(* IEC 61131-3 sources: IEC61131-3_ST_SCL_Mutation_Generator/Tests/mutatedCodeGenbit, 69 files *)

(* ---- M001.st ---- *)
FUNCTION_BLOCK GEN_BIT
  VAR_INPUT
    IN0 : DWORD;
    IN1 : DWORD;
    IN2 : DWORD;
    IN3 : DWORD;
    CLK : BOOL;
    STEPS : INT;
    REP : INT;
    RST : BOOL;
  END_VAR
  VAR_OUTPUT
    Q0 : BOOL;
    Q1 : BOOL;
    Q2 : BOOL;
    Q3 : BOOL;
    CNT : INT;
    RUN : BOOL;
  END_VAR
  VAR
    r0 : DWORD;
    r1 : DWORD;
    r2 : DWORD;
    r3 : DWORD;
    rx : INT := 1;
  END_VAR

  (* check if number of runs is finished or rep <> 0 which means continuous *) (* MUTATED: REL_OP_REPLACE *)

  IF clk AND NOT rst THEN
  	run := (rep = 0) OR (rx <= rep);
  	IF run THEN
  		(* check for step counter reached and reset to 0 if cnt = steps *)
  		IF cnt = steps THEN
  			cnt := 0;
  		END_IF;

  		(* when cnt = 0 then reload the inputs into the registers *)
  		IF cnt = 0 THEN
  			r0 := in0;
  			r1 := in1;
  			r2 := in2;
  			r3 := in3;
  		END_IF;

  		(* when cnt < steps, shift the lowest bits to the outputs *)
  		IF (cnt < steps) THEN
              Q0 := BIT_OF_DWORD(r0,0); (* Q0 := r0.X0; *)
              Q1 := BIT_OF_DWORD(r1,0); (* Q1 := r1.X0; *)
              Q2 := BIT_OF_DWORD(r2,0); (* Q2 := r2.X0; *)
              Q3 := BIT_OF_DWORD(r3,0); (* Q3 := r3.X0; *)
  			r0 := SHR(r0,1);
  			r1 := SHR(r1,1);
  			r2 := SHR(r2,1);
  			r3 := SHR(r3,1);
  		END_IF;

  		(* increment the step counter *)
  		cnt := cnt +1;
  		IF (cnt = steps) AND (rep <> 0) THEN rx := rx +1; END_IF;
  		IF (rx > rep) AND (rep <> 0) THEN run := FALSE; END_IF;
  	END_IF;
  ELSE
  	IF rst THEN
  		run := FALSE;
  		Q0 := FALSE;
  		Q1 := FALSE;
  		Q2 := FALSE;
  		Q3 := FALSE;
  		r0 := DWORD#0;
  		r1 := DWORD#0;
  		r2 := DWORD#0;
  		r3 := DWORD#0;
  		cnt := 0;
  		rx := 1;
  	END_IF;
  END_IF;

  (*From OSCAT Library, www.oscat.de *)
END_FUNCTION_BLOCK

(* ---- M002.st ---- *)
FUNCTION_BLOCK GEN_BIT
  VAR_INPUT
    IN0 : DWORD;
    IN1 : DWORD;
    IN2 : DWORD;
    IN3 : DWORD;
    CLK : BOOL;
    STEPS : INT;
    REP : INT;
    RST : BOOL;
  END_VAR
  VAR_OUTPUT
    Q0 : BOOL;
    Q1 : BOOL;
    Q2 : BOOL;
    Q3 : BOOL;
    CNT : INT;
    RUN : BOOL;
  END_VAR
  VAR
    r0 : DWORD;
    r1 : DWORD;
    r2 : DWORD;
    r3 : DWORD;
    rx : INT := 1;
  END_VAR

  (* check if number of runs is finished or rep = 0 which means continuous *)

  IF clk AND NOT rst THEN
  	run := (rep <> 0) OR (rx <= rep); (* MUTATED: REL_OP_REPLACE *)
  	IF run THEN
  		(* check for step counter reached and reset to 0 if cnt = steps *)
  		IF cnt = steps THEN
  			cnt := 0;
  		END_IF;

  		(* when cnt = 0 then reload the inputs into the registers *)
  		IF cnt = 0 THEN
  			r0 := in0;
  			r1 := in1;
  			r2 := in2;
  			r3 := in3;
  		END_IF;

  		(* when cnt < steps, shift the lowest bits to the outputs *)
  		IF (cnt < steps) THEN
              Q0 := BIT_OF_DWORD(r0,0); (* Q0 := r0.X0; *)
              Q1 := BIT_OF_DWORD(r1,0); (* Q1 := r1.X0; *)
              Q2 := BIT_OF_DWORD(r2,0); (* Q2 := r2.X0; *)
              Q3 := BIT_OF_DWORD(r3,0); (* Q3 := r3.X0; *)
  			r0 := SHR(r0,1);
  			r1 := SHR(r1,1);
  			r2 := SHR(r2,1);
  			r3 := SHR(r3,1);
  		END_IF;

  		(* increment the step counter *)
  		cnt := cnt +1;
  		IF (cnt = steps) AND (rep <> 0) THEN rx := rx +1; END_IF;
  		IF (rx > rep) AND (rep <> 0) THEN run := FALSE; END_IF;
  	END_IF;
  ELSE
  	IF rst THEN
  		run := FALSE;
  		Q0 := FALSE;
  		Q1 := FALSE;
  		Q2 := FALSE;
  		Q3 := FALSE;
  		r0 := DWORD#0;
  		r1 := DWORD#0;
  		r2 := DWORD#0;
  		r3 := DWORD#0;
  		cnt := 0;
  		rx := 1;
  	END_IF;
  END_IF;

  (*From OSCAT Library, www.oscat.de *)
END_FUNCTION_BLOCK

(* ---- M003.st ---- *)
FUNCTION_BLOCK GEN_BIT
  VAR_INPUT
    IN0 : DWORD;
    IN1 : DWORD;
    IN2 : DWORD;
    IN3 : DWORD;
    CLK : BOOL;
    STEPS : INT;
    REP : INT;
    RST : BOOL;
  END_VAR
  VAR_OUTPUT
    Q0 : BOOL;
    Q1 : BOOL;
    Q2 : BOOL;
    Q3 : BOOL;
    CNT : INT;
    RUN : BOOL;
  END_VAR
  VAR
    r0 : DWORD;
    r1 : DWORD;
    r2 : DWORD;
    r3 : DWORD;
    rx : INT := 1;
  END_VAR

  (* check if number of runs is finished or rep = 0 which means continuous *)

  IF clk AND NOT rst THEN
  	run := (rep = 0) OR (rx >= rep); (* MUTATED: REL_OP_REPLACE *)
  	IF run THEN
  		(* check for step counter reached and reset to 0 if cnt = steps *)
  		IF cnt = steps THEN
  			cnt := 0;
  		END_IF;

  		(* when cnt = 0 then reload the inputs into the registers *)
  		IF cnt = 0 THEN
  			r0 := in0;
  			r1 := in1;
  			r2 := in2;
  			r3 := in3;
  		END_IF;

  		(* when cnt < steps, shift the lowest bits to the outputs *)
  		IF (cnt < steps) THEN
              Q0 := BIT_OF_DWORD(r0,0); (* Q0 := r0.X0; *)
              Q1 := BIT_OF_DWORD(r1,0); (* Q1 := r1.X0; *)
              Q2 := BIT_OF_DWORD(r2,0); (* Q2 := r2.X0; *)
              Q3 := BIT_OF_DWORD(r3,0); (* Q3 := r3.X0; *)
  			r0 := SHR(r0,1);
  			r1 := SHR(r1,1);
  			r2 := SHR(r2,1);
  			r3 := SHR(r3,1);
  		END_IF;

  		(* increment the step counter *)
  		cnt := cnt +1;
  		IF (cnt = steps) AND (rep <> 0) THEN rx := rx +1; END_IF;
  		IF (rx > rep) AND (rep <> 0) THEN run := FALSE; END_IF;
  	END_IF;
  ELSE
  	IF rst THEN
  		run := FALSE;
  		Q0 := FALSE;
  		Q1 := FALSE;
  		Q2 := FALSE;
  		Q3 := FALSE;
  		r0 := DWORD#0;
  		r1 := DWORD#0;
  		r2 := DWORD#0;
  		r3 := DWORD#0;
  		cnt := 0;
  		rx := 1;
  	END_IF;
  END_IF;

  (*From OSCAT Library, www.oscat.de *)
END_FUNCTION_BLOCK

(* ---- M004.st ---- *)
FUNCTION_BLOCK GEN_BIT
  VAR_INPUT
    IN0 : DWORD;
    IN1 : DWORD;
    IN2 : DWORD;
    IN3 : DWORD;
    CLK : BOOL;
    STEPS : INT;
    REP : INT;
    RST : BOOL;
  END_VAR
  VAR_OUTPUT
    Q0 : BOOL;
    Q1 : BOOL;
    Q2 : BOOL;
    Q3 : BOOL;
    CNT : INT;
    RUN : BOOL;
  END_VAR
  VAR
    r0 : DWORD;
    r1 : DWORD;
    r2 : DWORD;
    r3 : DWORD;
    rx : INT := 1;
  END_VAR

  (* check if number of runs is finished or rep = 0 which means continuous *)

  IF clk AND NOT rst THEN
  	run := (rep = 0) OR (rx <= rep);
  	IF run THEN
  		(* check for step counter reached and reset to 0 if cnt <> steps *) (* MUTATED: REL_OP_REPLACE *)
  		IF cnt = steps THEN
  			cnt := 0;
  		END_IF;

  		(* when cnt = 0 then reload the inputs into the registers *)
  		IF cnt = 0 THEN
  			r0 := in0;
  			r1 := in1;
  			r2 := in2;
  			r3 := in3;
  		END_IF;

  		(* when cnt < steps, shift the lowest bits to the outputs *)
  		IF (cnt < steps) THEN
              Q0 := BIT_OF_DWORD(r0,0); (* Q0 := r0.X0; *)
              Q1 := BIT_OF_DWORD(r1,0); (* Q1 := r1.X0; *)
              Q2 := BIT_OF_DWORD(r2,0); (* Q2 := r2.X0; *)
              Q3 := BIT_OF_DWORD(r3,0); (* Q3 := r3.X0; *)
  			r0 := SHR(r0,1);
  			r1 := SHR(r1,1);
  			r2 := SHR(r2,1);
  			r3 := SHR(r3,1);
  		END_IF;

  		(* increment the step counter *)
  		cnt := cnt +1;
  		IF (cnt = steps) AND (rep <> 0) THEN rx := rx +1; END_IF;
  		IF (rx > rep) AND (rep <> 0) THEN run := FALSE; END_IF;
  	END_IF;
  ELSE
  	IF rst THEN
  		run := FALSE;
  		Q0 := FALSE;
  		Q1 := FALSE;
  		Q2 := FALSE;
  		Q3 := FALSE;
  		r0 := DWORD#0;
  		r1 := DWORD#0;
  		r2 := DWORD#0;
  		r3 := DWORD#0;
  		cnt := 0;
  		rx := 1;
  	END_IF;
  END_IF;

  (*From OSCAT Library, www.oscat.de *)
END_FUNCTION_BLOCK

(* ---- M005.st ---- *)
FUNCTION_BLOCK GEN_BIT
  VAR_INPUT
    IN0 : DWORD;
    IN1 : DWORD;
    IN2 : DWORD;
    IN3 : DWORD;
    CLK : BOOL;
    STEPS : INT;
    REP : INT;
    RST : BOOL;
  END_VAR
  VAR_OUTPUT
    Q0 : BOOL;
    Q1 : BOOL;
    Q2 : BOOL;
    Q3 : BOOL;
    CNT : INT;
    RUN : BOOL;
  END_VAR
  VAR
    r0 : DWORD;
    r1 : DWORD;
    r2 : DWORD;
    r3 : DWORD;
    rx : INT := 1;
  END_VAR

  (* check if number of runs is finished or rep = 0 which means continuous *)

  IF clk AND NOT rst THEN
  	run := (rep = 0) OR (rx <= rep);
  	IF run THEN
  		(* check for step counter reached and reset to 0 if cnt = steps *)
  		IF cnt <> steps THEN (* MUTATED: REL_OP_REPLACE *)
  			cnt := 0;
  		END_IF;

  		(* when cnt = 0 then reload the inputs into the registers *)
  		IF cnt = 0 THEN
  			r0 := in0;
  			r1 := in1;
  			r2 := in2;
  			r3 := in3;
  		END_IF;

  		(* when cnt < steps, shift the lowest bits to the outputs *)
  		IF (cnt < steps) THEN
              Q0 := BIT_OF_DWORD(r0,0); (* Q0 := r0.X0; *)
              Q1 := BIT_OF_DWORD(r1,0); (* Q1 := r1.X0; *)
              Q2 := BIT_OF_DWORD(r2,0); (* Q2 := r2.X0; *)
              Q3 := BIT_OF_DWORD(r3,0); (* Q3 := r3.X0; *)
  			r0 := SHR(r0,1);
  			r1 := SHR(r1,1);
  			r2 := SHR(r2,1);
  			r3 := SHR(r3,1);
  		END_IF;

  		(* increment the step counter *)
  		cnt := cnt +1;
  		IF (cnt = steps) AND (rep <> 0) THEN rx := rx +1; END_IF;
  		IF (rx > rep) AND (rep <> 0) THEN run := FALSE; END_IF;
  	END_IF;
  ELSE
  	IF rst THEN
  		run := FALSE;
  		Q0 := FALSE;
  		Q1 := FALSE;
  		Q2 := FALSE;
  		Q3 := FALSE;
  		r0 := DWORD#0;
  		r1 := DWORD#0;
  		r2 := DWORD#0;
  		r3 := DWORD#0;
  		cnt := 0;
  		rx := 1;
  	END_IF;
  END_IF;

  (*From OSCAT Library, www.oscat.de *)
END_FUNCTION_BLOCK

(* ---- M006.st ---- *)
FUNCTION_BLOCK GEN_BIT
  VAR_INPUT
    IN0 : DWORD;
    IN1 : DWORD;
    IN2 : DWORD;
    IN3 : DWORD;
    CLK : BOOL;
    STEPS : INT;
    REP : INT;
    RST : BOOL;
  END_VAR
  VAR_OUTPUT
    Q0 : BOOL;
    Q1 : BOOL;
    Q2 : BOOL;
    Q3 : BOOL;
    CNT : INT;
    RUN : BOOL;
  END_VAR
  VAR
    r0 : DWORD;
    r1 : DWORD;
    r2 : DWORD;
    r3 : DWORD;
    rx : INT := 1;
  END_VAR

  (* check if number of runs is finished or rep = 0 which means continuous *)

  IF clk AND NOT rst THEN
  	run := (rep = 0) OR (rx <= rep);
  	IF run THEN
  		(* check for step counter reached and reset to 0 if cnt = steps *)
  		IF cnt = steps THEN
  			cnt := 0;
  		END_IF;

  		(* when cnt <> 0 then reload the inputs into the registers *) (* MUTATED: REL_OP_REPLACE *)
  		IF cnt = 0 THEN
  			r0 := in0;
  			r1 := in1;
  			r2 := in2;
  			r3 := in3;
  		END_IF;

  		(* when cnt < steps, shift the lowest bits to the outputs *)
  		IF (cnt < steps) THEN
              Q0 := BIT_OF_DWORD(r0,0); (* Q0 := r0.X0; *)
              Q1 := BIT_OF_DWORD(r1,0); (* Q1 := r1.X0; *)
              Q2 := BIT_OF_DWORD(r2,0); (* Q2 := r2.X0; *)
              Q3 := BIT_OF_DWORD(r3,0); (* Q3 := r3.X0; *)
  			r0 := SHR(r0,1);
  			r1 := SHR(r1,1);
  			r2 := SHR(r2,1);
  			r3 := SHR(r3,1);
  		END_IF;

  		(* increment the step counter *)
  		cnt := cnt +1;
  		IF (cnt = steps) AND (rep <> 0) THEN rx := rx +1; END_IF;
  		IF (rx > rep) AND (rep <> 0) THEN run := FALSE; END_IF;
  	END_IF;
  ELSE
  	IF rst THEN
  		run := FALSE;
  		Q0 := FALSE;
  		Q1 := FALSE;
  		Q2 := FALSE;
  		Q3 := FALSE;
  		r0 := DWORD#0;
  		r1 := DWORD#0;
  		r2 := DWORD#0;
  		r3 := DWORD#0;
  		cnt := 0;
  		rx := 1;
  	END_IF;
  END_IF;

  (*From OSCAT Library, www.oscat.de *)
END_FUNCTION_BLOCK

(* ---- M007.st ---- *)
FUNCTION_BLOCK GEN_BIT
  VAR_INPUT
    IN0 : DWORD;
    IN1 : DWORD;
    IN2 : DWORD;
    IN3 : DWORD;
    CLK : BOOL;
    STEPS : INT;
    REP : INT;
    RST : BOOL;
  END_VAR
  VAR_OUTPUT
    Q0 : BOOL;
    Q1 : BOOL;
    Q2 : BOOL;
    Q3 : BOOL;
    CNT : INT;
    RUN : BOOL;
  END_VAR
  VAR
    r0 : DWORD;
    r1 : DWORD;
    r2 : DWORD;
    r3 : DWORD;
    rx : INT := 1;
  END_VAR

  (* check if number of runs is finished or rep = 0 which means continuous *)

  IF clk AND NOT rst THEN
  	run := (rep = 0) OR (rx <= rep);
  	IF run THEN
  		(* check for step counter reached and reset to 0 if cnt = steps *)
  		IF cnt = steps THEN
  			cnt := 0;
  		END_IF;

  		(* when cnt = 0 then reload the inputs into the registers *)
  		IF cnt <> 0 THEN (* MUTATED: REL_OP_REPLACE *)
  			r0 := in0;
  			r1 := in1;
  			r2 := in2;
  			r3 := in3;
  		END_IF;

  		(* when cnt < steps, shift the lowest bits to the outputs *)
  		IF (cnt < steps) THEN
              Q0 := BIT_OF_DWORD(r0,0); (* Q0 := r0.X0; *)
              Q1 := BIT_OF_DWORD(r1,0); (* Q1 := r1.X0; *)
              Q2 := BIT_OF_DWORD(r2,0); (* Q2 := r2.X0; *)
              Q3 := BIT_OF_DWORD(r3,0); (* Q3 := r3.X0; *)
  			r0 := SHR(r0,1);
  			r1 := SHR(r1,1);
  			r2 := SHR(r2,1);
  			r3 := SHR(r3,1);
  		END_IF;

  		(* increment the step counter *)
  		cnt := cnt +1;
  		IF (cnt = steps) AND (rep <> 0) THEN rx := rx +1; END_IF;
  		IF (rx > rep) AND (rep <> 0) THEN run := FALSE; END_IF;
  	END_IF;
  ELSE
  	IF rst THEN
  		run := FALSE;
  		Q0 := FALSE;
  		Q1 := FALSE;
  		Q2 := FALSE;
  		Q3 := FALSE;
  		r0 := DWORD#0;
  		r1 := DWORD#0;
  		r2 := DWORD#0;
  		r3 := DWORD#0;
  		cnt := 0;
  		rx := 1;
  	END_IF;
  END_IF;

  (*From OSCAT Library, www.oscat.de *)
END_FUNCTION_BLOCK

(* ---- M008.st ---- *)
FUNCTION_BLOCK GEN_BIT
  VAR_INPUT
    IN0 : DWORD;
    IN1 : DWORD;
    IN2 : DWORD;
    IN3 : DWORD;
    CLK : BOOL;
    STEPS : INT;
    REP : INT;
    RST : BOOL;
  END_VAR
  VAR_OUTPUT
    Q0 : BOOL;
    Q1 : BOOL;
    Q2 : BOOL;
    Q3 : BOOL;
    CNT : INT;
    RUN : BOOL;
  END_VAR
  VAR
    r0 : DWORD;
    r1 : DWORD;
    r2 : DWORD;
    r3 : DWORD;
    rx : INT := 1;
  END_VAR

  (* check if number of runs is finished or rep = 0 which means continuous *)

  IF clk AND NOT rst THEN
  	run := (rep = 0) OR (rx <= rep);
  	IF run THEN
  		(* check for step counter reached and reset to 0 if cnt = steps *)
  		IF cnt = steps THEN
  			cnt := 0;
  		END_IF;

  		(* when cnt = 0 then reload the inputs into the registers *)
  		IF cnt = 0 THEN
  			r0 := in0;
  			r1 := in1;
  			r2 := in2;
  			r3 := in3;
  		END_IF;

  		(* when cnt > steps, shift the lowest bits to the outputs *) (* MUTATED: REL_OP_REPLACE *)
  		IF (cnt < steps) THEN
              Q0 := BIT_OF_DWORD(r0,0); (* Q0 := r0.X0; *)
              Q1 := BIT_OF_DWORD(r1,0); (* Q1 := r1.X0; *)
              Q2 := BIT_OF_DWORD(r2,0); (* Q2 := r2.X0; *)
              Q3 := BIT_OF_DWORD(r3,0); (* Q3 := r3.X0; *)
  			r0 := SHR(r0,1);
  			r1 := SHR(r1,1);
  			r2 := SHR(r2,1);
  			r3 := SHR(r3,1);
  		END_IF;

  		(* increment the step counter *)
  		cnt := cnt +1;
  		IF (cnt = steps) AND (rep <> 0) THEN rx := rx +1; END_IF;
  		IF (rx > rep) AND (rep <> 0) THEN run := FALSE; END_IF;
  	END_IF;
  ELSE
  	IF rst THEN
  		run := FALSE;
  		Q0 := FALSE;
  		Q1 := FALSE;
  		Q2 := FALSE;
  		Q3 := FALSE;
  		r0 := DWORD#0;
  		r1 := DWORD#0;
  		r2 := DWORD#0;
  		r3 := DWORD#0;
  		cnt := 0;
  		rx := 1;
  	END_IF;
  END_IF;

  (*From OSCAT Library, www.oscat.de *)
END_FUNCTION_BLOCK

(* ---- M009.st ---- *)
FUNCTION_BLOCK GEN_BIT
  VAR_INPUT
    IN0 : DWORD;
    IN1 : DWORD;
    IN2 : DWORD;
    IN3 : DWORD;
    CLK : BOOL;
    STEPS : INT;
    REP : INT;
    RST : BOOL;
  END_VAR
  VAR_OUTPUT
    Q0 : BOOL;
    Q1 : BOOL;
    Q2 : BOOL;
    Q3 : BOOL;
    CNT : INT;
    RUN : BOOL;
  END_VAR
  VAR
    r0 : DWORD;
    r1 : DWORD;
    r2 : DWORD;
    r3 : DWORD;
    rx : INT := 1;
  END_VAR

  (* check if number of runs is finished or rep = 0 which means continuous *)

  IF clk AND NOT rst THEN
  	run := (rep = 0) OR (rx <= rep);
  	IF run THEN
  		(* check for step counter reached and reset to 0 if cnt = steps *)
  		IF cnt = steps THEN
  			cnt := 0;
  		END_IF;

  		(* when cnt = 0 then reload the inputs into the registers *)
  		IF cnt = 0 THEN
  			r0 := in0;
  			r1 := in1;
  			r2 := in2;
  			r3 := in3;
  		END_IF;

  		(* when cnt < steps, shift the lowest bits to the outputs *)
  		IF (cnt > steps) THEN (* MUTATED: REL_OP_REPLACE *)
              Q0 := BIT_OF_DWORD(r0,0); (* Q0 := r0.X0; *)
              Q1 := BIT_OF_DWORD(r1,0); (* Q1 := r1.X0; *)
              Q2 := BIT_OF_DWORD(r2,0); (* Q2 := r2.X0; *)
              Q3 := BIT_OF_DWORD(r3,0); (* Q3 := r3.X0; *)
  			r0 := SHR(r0,1);
  			r1 := SHR(r1,1);
  			r2 := SHR(r2,1);
  			r3 := SHR(r3,1);
  		END_IF;

  		(* increment the step counter *)
  		cnt := cnt +1;
  		IF (cnt = steps) AND (rep <> 0) THEN rx := rx +1; END_IF;
  		IF (rx > rep) AND (rep <> 0) THEN run := FALSE; END_IF;
  	END_IF;
  ELSE
  	IF rst THEN
  		run := FALSE;
  		Q0 := FALSE;
  		Q1 := FALSE;
  		Q2 := FALSE;
  		Q3 := FALSE;
  		r0 := DWORD#0;
  		r1 := DWORD#0;
  		r2 := DWORD#0;
  		r3 := DWORD#0;
  		cnt := 0;
  		rx := 1;
  	END_IF;
  END_IF;

  (*From OSCAT Library, www.oscat.de *)
END_FUNCTION_BLOCK

(* ---- M010.st ---- *)
FUNCTION_BLOCK GEN_BIT
  VAR_INPUT
    IN0 : DWORD;
    IN1 : DWORD;
    IN2 : DWORD;
    IN3 : DWORD;
    CLK : BOOL;
    STEPS : INT;
    REP : INT;
    RST : BOOL;
  END_VAR
  VAR_OUTPUT
    Q0 : BOOL;
    Q1 : BOOL;
    Q2 : BOOL;
    Q3 : BOOL;
    CNT : INT;
    RUN : BOOL;
  END_VAR
  VAR
    r0 : DWORD;
    r1 : DWORD;
    r2 : DWORD;
    r3 : DWORD;
    rx : INT := 1;
  END_VAR

  (* check if number of runs is finished or rep = 0 which means continuous *)

  IF clk AND NOT rst THEN
  	run := (rep = 0) OR (rx <= rep);
  	IF run THEN
  		(* check for step counter reached and reset to 0 if cnt = steps *)
  		IF cnt = steps THEN
  			cnt := 0;
  		END_IF;

  		(* when cnt = 0 then reload the inputs into the registers *)
  		IF cnt = 0 THEN
  			r0 := in0;
  			r1 := in1;
  			r2 := in2;
  			r3 := in3;
  		END_IF;

  		(* when cnt < steps, shift the lowest bits to the outputs *)
  		IF (cnt < steps) THEN
              Q0 := BIT_OF_DWORD(r0,0); (* Q0 := r0.X0; *)
              Q1 := BIT_OF_DWORD(r1,0); (* Q1 := r1.X0; *)
              Q2 := BIT_OF_DWORD(r2,0); (* Q2 := r2.X0; *)
              Q3 := BIT_OF_DWORD(r3,0); (* Q3 := r3.X0; *)
  			r0 := SHR(r0,1);
  			r1 := SHR(r1,1);
  			r2 := SHR(r2,1);
  			r3 := SHR(r3,1);
  		END_IF;

  		(* increment the step counter *)
  		cnt := cnt +1;
  		IF (cnt <> steps) AND (rep <> 0) THEN rx := rx +1; END_IF; (* MUTATED: REL_OP_REPLACE *)
  		IF (rx > rep) AND (rep <> 0) THEN run := FALSE; END_IF;
  	END_IF;
  ELSE
  	IF rst THEN
  		run := FALSE;
  		Q0 := FALSE;
  		Q1 := FALSE;
  		Q2 := FALSE;
  		Q3 := FALSE;
  		r0 := DWORD#0;
  		r1 := DWORD#0;
  		r2 := DWORD#0;
  		r3 := DWORD#0;
  		cnt := 0;
  		rx := 1;
  	END_IF;
  END_IF;

  (*From OSCAT Library, www.oscat.de *)
END_FUNCTION_BLOCK

(* ---- M011.st ---- *)
FUNCTION_BLOCK GEN_BIT
  VAR_INPUT
    IN0 : DWORD;
    IN1 : DWORD;
    IN2 : DWORD;
    IN3 : DWORD;
    CLK : BOOL;
    STEPS : INT;
    REP : INT;
    RST : BOOL;
  END_VAR
  VAR_OUTPUT
    Q0 : BOOL;
    Q1 : BOOL;
    Q2 : BOOL;
    Q3 : BOOL;
    CNT : INT;
    RUN : BOOL;
  END_VAR
  VAR
    r0 : DWORD;
    r1 : DWORD;
    r2 : DWORD;
    r3 : DWORD;
    rx : INT := 1;
  END_VAR

  (* check if number of runs is finished or rep = 0 which means continuous *)

  IF clk AND NOT rst THEN
  	run := (rep = 0) OR (rx <= rep);
  	IF run THEN
  		(* check for step counter reached and reset to 0 if cnt = steps *)
  		IF cnt = steps THEN
  			cnt := 0;
  		END_IF;

  		(* when cnt = 0 then reload the inputs into the registers *)
  		IF cnt = 0 THEN
  			r0 := in0;
  			r1 := in1;
  			r2 := in2;
  			r3 := in3;
  		END_IF;

  		(* when cnt < steps, shift the lowest bits to the outputs *)
  		IF (cnt < steps) THEN
              Q0 := BIT_OF_DWORD(r0,0); (* Q0 := r0.X0; *)
              Q1 := BIT_OF_DWORD(r1,0); (* Q1 := r1.X0; *)
              Q2 := BIT_OF_DWORD(r2,0); (* Q2 := r2.X0; *)
              Q3 := BIT_OF_DWORD(r3,0); (* Q3 := r3.X0; *)
  			r0 := SHR(r0,1);
  			r1 := SHR(r1,1);
  			r2 := SHR(r2,1);
  			r3 := SHR(r3,1);
  		END_IF;

  		(* increment the step counter *)
  		cnt := cnt +1;
  		IF (cnt = steps) AND (rep = 0) THEN rx := rx +1; END_IF; (* MUTATED: REL_OP_REPLACE *)
  		IF (rx > rep) AND (rep <> 0) THEN run := FALSE; END_IF;
  	END_IF;
  ELSE
  	IF rst THEN
  		run := FALSE;
  		Q0 := FALSE;
  		Q1 := FALSE;
  		Q2 := FALSE;
  		Q3 := FALSE;
  		r0 := DWORD#0;
  		r1 := DWORD#0;
  		r2 := DWORD#0;
  		r3 := DWORD#0;
  		cnt := 0;
  		rx := 1;
  	END_IF;
  END_IF;

  (*From OSCAT Library, www.oscat.de *)
END_FUNCTION_BLOCK

(* ---- M012.st ---- *)
FUNCTION_BLOCK GEN_BIT
  VAR_INPUT
    IN0 : DWORD;
    IN1 : DWORD;
    IN2 : DWORD;
    IN3 : DWORD;
    CLK : BOOL;
    STEPS : INT;
    REP : INT;
    RST : BOOL;
  END_VAR
  VAR_OUTPUT
    Q0 : BOOL;
    Q1 : BOOL;
    Q2 : BOOL;
    Q3 : BOOL;
    CNT : INT;
    RUN : BOOL;
  END_VAR
  VAR
    r0 : DWORD;
    r1 : DWORD;
    r2 : DWORD;
    r3 : DWORD;
    rx : INT := 1;
  END_VAR

  (* check if number of runs is finished or rep = 0 which means continuous *)

  IF clk AND NOT rst THEN
  	run := (rep = 0) OR (rx <= rep);
  	IF run THEN
  		(* check for step counter reached and reset to 0 if cnt = steps *)
  		IF cnt = steps THEN
  			cnt := 0;
  		END_IF;

  		(* when cnt = 0 then reload the inputs into the registers *)
  		IF cnt = 0 THEN
  			r0 := in0;
  			r1 := in1;
  			r2 := in2;
  			r3 := in3;
  		END_IF;

  		(* when cnt < steps, shift the lowest bits to the outputs *)
  		IF (cnt < steps) THEN
              Q0 := BIT_OF_DWORD(r0,0); (* Q0 := r0.X0; *)
              Q1 := BIT_OF_DWORD(r1,0); (* Q1 := r1.X0; *)
              Q2 := BIT_OF_DWORD(r2,0); (* Q2 := r2.X0; *)
              Q3 := BIT_OF_DWORD(r3,0); (* Q3 := r3.X0; *)
  			r0 := SHR(r0,1);
  			r1 := SHR(r1,1);
  			r2 := SHR(r2,1);
  			r3 := SHR(r3,1);
  		END_IF;

  		(* increment the step counter *)
  		cnt := cnt +1;
  		IF (cnt = steps) AND (rep <> 0) THEN rx := rx +1; END_IF;
  		IF (rx < rep) AND (rep <> 0) THEN run := FALSE; END_IF; (* MUTATED: REL_OP_REPLACE *)
  	END_IF;
  ELSE
  	IF rst THEN
  		run := FALSE;
  		Q0 := FALSE;
  		Q1 := FALSE;
  		Q2 := FALSE;
  		Q3 := FALSE;
  		r0 := DWORD#0;
  		r1 := DWORD#0;
  		r2 := DWORD#0;
  		r3 := DWORD#0;
  		cnt := 0;
  		rx := 1;
  	END_IF;
  END_IF;

  (*From OSCAT Library, www.oscat.de *)
END_FUNCTION_BLOCK

(* ---- M013.st ---- *)
FUNCTION_BLOCK GEN_BIT
  VAR_INPUT
    IN0 : DWORD;
    IN1 : DWORD;
    IN2 : DWORD;
    IN3 : DWORD;
    CLK : BOOL;
    STEPS : INT;
    REP : INT;
    RST : BOOL;
  END_VAR
  VAR_OUTPUT
    Q0 : BOOL;
    Q1 : BOOL;
    Q2 : BOOL;
    Q3 : BOOL;
    CNT : INT;
    RUN : BOOL;
  END_VAR
  VAR
    r0 : DWORD;
    r1 : DWORD;
    r2 : DWORD;
    r3 : DWORD;
    rx : INT := 1;
  END_VAR

  (* check if number of runs is finished or rep = 0 which means continuous *)

  IF clk AND NOT rst THEN
  	run := (rep = 0) OR (rx <= rep);
  	IF run THEN
  		(* check for step counter reached and reset to 0 if cnt = steps *)
  		IF cnt = steps THEN
  			cnt := 0;
  		END_IF;

  		(* when cnt = 0 then reload the inputs into the registers *)
  		IF cnt = 0 THEN
  			r0 := in0;
  			r1 := in1;
  			r2 := in2;
  			r3 := in3;
  		END_IF;

  		(* when cnt < steps, shift the lowest bits to the outputs *)
  		IF (cnt < steps) THEN
              Q0 := BIT_OF_DWORD(r0,0); (* Q0 := r0.X0; *)
              Q1 := BIT_OF_DWORD(r1,0); (* Q1 := r1.X0; *)
              Q2 := BIT_OF_DWORD(r2,0); (* Q2 := r2.X0; *)
              Q3 := BIT_OF_DWORD(r3,0); (* Q3 := r3.X0; *)
  			r0 := SHR(r0,1);
  			r1 := SHR(r1,1);
  			r2 := SHR(r2,1);
  			r3 := SHR(r3,1);
  		END_IF;

  		(* increment the step counter *)
  		cnt := cnt +1;
  		IF (cnt = steps) AND (rep <> 0) THEN rx := rx +1; END_IF;
  		IF (rx > rep) AND (rep = 0) THEN run := FALSE; END_IF; (* MUTATED: REL_OP_REPLACE *)
  	END_IF;
  ELSE
  	IF rst THEN
  		run := FALSE;
  		Q0 := FALSE;
  		Q1 := FALSE;
  		Q2 := FALSE;
  		Q3 := FALSE;
  		r0 := DWORD#0;
  		r1 := DWORD#0;
  		r2 := DWORD#0;
  		r3 := DWORD#0;
  		cnt := 0;
  		rx := 1;
  	END_IF;
  END_IF;

  (*From OSCAT Library, www.oscat.de *)
END_FUNCTION_BLOCK

(* ---- M014.st ---- *)
FUNCTION_BLOCK GEN_BIT
  VAR_INPUT
    IN0 : DWORD;
    IN1 : DWORD;
    IN2 : DWORD;
    IN3 : DWORD;
    CLK : BOOL;
    STEPS : INT;
    REP : INT;
    RST : BOOL;
  END_VAR
  VAR_OUTPUT
    Q0 : BOOL;
    Q1 : BOOL;
    Q2 : BOOL;
    Q3 : BOOL;
    CNT : INT;
    RUN : BOOL;
  END_VAR
  VAR
    r0 : DWORD;
    r1 : DWORD;
    r2 : DWORD;
    r3 : DWORD;
    rx : INT := 1;
  END_VAR

  (* check if number of runs is finished or rep = 0 which means continuous *)

  IF clk OR NOT rst THEN (* MUTATED: LOGICAL_OP_REPLACE *)
  	run := (rep = 0) OR (rx <= rep);
  	IF run THEN
  		(* check for step counter reached and reset to 0 if cnt = steps *)
  		IF cnt = steps THEN
  			cnt := 0;
  		END_IF;

  		(* when cnt = 0 then reload the inputs into the registers *)
  		IF cnt = 0 THEN
  			r0 := in0;
  			r1 := in1;
  			r2 := in2;
  			r3 := in3;
  		END_IF;

  		(* when cnt < steps, shift the lowest bits to the outputs *)
  		IF (cnt < steps) THEN
              Q0 := BIT_OF_DWORD(r0,0); (* Q0 := r0.X0; *)
              Q1 := BIT_OF_DWORD(r1,0); (* Q1 := r1.X0; *)
              Q2 := BIT_OF_DWORD(r2,0); (* Q2 := r2.X0; *)
              Q3 := BIT_OF_DWORD(r3,0); (* Q3 := r3.X0; *)
  			r0 := SHR(r0,1);
  			r1 := SHR(r1,1);
  			r2 := SHR(r2,1);
  			r3 := SHR(r3,1);
  		END_IF;

  		(* increment the step counter *)
  		cnt := cnt +1;
  		IF (cnt = steps) AND (rep <> 0) THEN rx := rx +1; END_IF;
  		IF (rx > rep) AND (rep <> 0) THEN run := FALSE; END_IF;
  	END_IF;
  ELSE
  	IF rst THEN
  		run := FALSE;
  		Q0 := FALSE;
  		Q1 := FALSE;
  		Q2 := FALSE;
  		Q3 := FALSE;
  		r0 := DWORD#0;
  		r1 := DWORD#0;
  		r2 := DWORD#0;
  		r3 := DWORD#0;
  		cnt := 0;
  		rx := 1;
  	END_IF;
  END_IF;

  (*From OSCAT Library, www.oscat.de *)
END_FUNCTION_BLOCK

(* ---- M015.st ---- *)
FUNCTION_BLOCK GEN_BIT
  VAR_INPUT
    IN0 : DWORD;
    IN1 : DWORD;
    IN2 : DWORD;
    IN3 : DWORD;
    CLK : BOOL;
    STEPS : INT;
    REP : INT;
    RST : BOOL;
  END_VAR
  VAR_OUTPUT
    Q0 : BOOL;
    Q1 : BOOL;
    Q2 : BOOL;
    Q3 : BOOL;
    CNT : INT;
    RUN : BOOL;
  END_VAR
  VAR
    r0 : DWORD;
    r1 : DWORD;
    r2 : DWORD;
    r3 : DWORD;
    rx : INT := 1;
  END_VAR

  (* check if number of runs is finished or rep = 0 which means continuous *)

  IF clk AND NOT rst THEN
  	run := (rep = 0) AND (rx <= rep); (* MUTATED: LOGICAL_OP_REPLACE *)
  	IF run THEN
  		(* check for step counter reached and reset to 0 if cnt = steps *)
  		IF cnt = steps THEN
  			cnt := 0;
  		END_IF;

  		(* when cnt = 0 then reload the inputs into the registers *)
  		IF cnt = 0 THEN
  			r0 := in0;
  			r1 := in1;
  			r2 := in2;
  			r3 := in3;
  		END_IF;

  		(* when cnt < steps, shift the lowest bits to the outputs *)
  		IF (cnt < steps) THEN
              Q0 := BIT_OF_DWORD(r0,0); (* Q0 := r0.X0; *)
              Q1 := BIT_OF_DWORD(r1,0); (* Q1 := r1.X0; *)
              Q2 := BIT_OF_DWORD(r2,0); (* Q2 := r2.X0; *)
              Q3 := BIT_OF_DWORD(r3,0); (* Q3 := r3.X0; *)
  			r0 := SHR(r0,1);
  			r1 := SHR(r1,1);
  			r2 := SHR(r2,1);
  			r3 := SHR(r3,1);
  		END_IF;

  		(* increment the step counter *)
  		cnt := cnt +1;
  		IF (cnt = steps) AND (rep <> 0) THEN rx := rx +1; END_IF;
  		IF (rx > rep) AND (rep <> 0) THEN run := FALSE; END_IF;
  	END_IF;
  ELSE
  	IF rst THEN
  		run := FALSE;
  		Q0 := FALSE;
  		Q1 := FALSE;
  		Q2 := FALSE;
  		Q3 := FALSE;
  		r0 := DWORD#0;
  		r1 := DWORD#0;
  		r2 := DWORD#0;
  		r3 := DWORD#0;
  		cnt := 0;
  		rx := 1;
  	END_IF;
  END_IF;

  (*From OSCAT Library, www.oscat.de *)
END_FUNCTION_BLOCK

(* ---- M016.st ---- *)
FUNCTION_BLOCK GEN_BIT
  VAR_INPUT
    IN0 : DWORD;
    IN1 : DWORD;
    IN2 : DWORD;
    IN3 : DWORD;
    CLK : BOOL;
    STEPS : INT;
    REP : INT;
    RST : BOOL;
  END_VAR
  VAR_OUTPUT
    Q0 : BOOL;
    Q1 : BOOL;
    Q2 : BOOL;
    Q3 : BOOL;
    CNT : INT;
    RUN : BOOL;
  END_VAR
  VAR
    r0 : DWORD;
    r1 : DWORD;
    r2 : DWORD;
    r3 : DWORD;
    rx : INT := 1;
  END_VAR

  (* check if number of runs is finished or rep = 0 which means continuous *)

  IF clk AND NOT rst THEN
  	run := (rep = 0) OR (rx <= rep);
  	IF run THEN
  		(* check for step counter reached and reset to 0 if cnt = steps *)
  		IF cnt = steps THEN
  			cnt := 0;
  		END_IF;

  		(* when cnt = 0 then reload the inputs into the registers *)
  		IF cnt = 0 THEN
  			r0 := in0;
  			r1 := in1;
  			r2 := in2;
  			r3 := in3;
  		END_IF;

  		(* when cnt < steps, shift the lowest bits to the outputs *)
  		IF (cnt < steps) THEN
              Q0 := BIT_OF_DWORD(r0,0); (* Q0 := r0.X0; *)
              Q1 := BIT_OF_DWORD(r1,0); (* Q1 := r1.X0; *)
              Q2 := BIT_OF_DWORD(r2,0); (* Q2 := r2.X0; *)
              Q3 := BIT_OF_DWORD(r3,0); (* Q3 := r3.X0; *)
  			r0 := SHR(r0,1);
  			r1 := SHR(r1,1);
  			r2 := SHR(r2,1);
  			r3 := SHR(r3,1);
  		END_IF;

  		(* increment the step counter *)
  		cnt := cnt +1;
  		IF (cnt = steps) OR (rep <> 0) THEN rx := rx +1; END_IF; (* MUTATED: LOGICAL_OP_REPLACE *)
  		IF (rx > rep) AND (rep <> 0) THEN run := FALSE; END_IF;
  	END_IF;
  ELSE
  	IF rst THEN
  		run := FALSE;
  		Q0 := FALSE;
  		Q1 := FALSE;
  		Q2 := FALSE;
  		Q3 := FALSE;
  		r0 := DWORD#0;
  		r1 := DWORD#0;
  		r2 := DWORD#0;
  		r3 := DWORD#0;
  		cnt := 0;
  		rx := 1;
  	END_IF;
  END_IF;

  (*From OSCAT Library, www.oscat.de *)
END_FUNCTION_BLOCK

(* ---- M017.st ---- *)
FUNCTION_BLOCK GEN_BIT
  VAR_INPUT
    IN0 : DWORD;
    IN1 : DWORD;
    IN2 : DWORD;
    IN3 : DWORD;
    CLK : BOOL;
    STEPS : INT;
    REP : INT;
    RST : BOOL;
  END_VAR
  VAR_OUTPUT
    Q0 : BOOL;
    Q1 : BOOL;
    Q2 : BOOL;
    Q3 : BOOL;
    CNT : INT;
    RUN : BOOL;
  END_VAR
  VAR
    r0 : DWORD;
    r1 : DWORD;
    r2 : DWORD;
    r3 : DWORD;
    rx : INT := 1;
  END_VAR

  (* check if number of runs is finished or rep = 0 which means continuous *)

  IF clk AND NOT rst THEN
  	run := (rep = 0) OR (rx <= rep);
  	IF run THEN
  		(* check for step counter reached and reset to 0 if cnt = steps *)
  		IF cnt = steps THEN
  			cnt := 0;
  		END_IF;

  		(* when cnt = 0 then reload the inputs into the registers *)
  		IF cnt = 0 THEN
  			r0 := in0;
  			r1 := in1;
  			r2 := in2;
  			r3 := in3;
  		END_IF;

  		(* when cnt < steps, shift the lowest bits to the outputs *)
  		IF (cnt < steps) THEN
              Q0 := BIT_OF_DWORD(r0,0); (* Q0 := r0.X0; *)
              Q1 := BIT_OF_DWORD(r1,0); (* Q1 := r1.X0; *)
              Q2 := BIT_OF_DWORD(r2,0); (* Q2 := r2.X0; *)
              Q3 := BIT_OF_DWORD(r3,0); (* Q3 := r3.X0; *)
  			r0 := SHR(r0,1);
  			r1 := SHR(r1,1);
  			r2 := SHR(r2,1);
  			r3 := SHR(r3,1);
  		END_IF;

  		(* increment the step counter *)
  		cnt := cnt +1;
  		IF (cnt = steps) AND (rep <> 0) THEN rx := rx +1; END_IF;
  		IF (rx > rep) OR (rep <> 0) THEN run := FALSE; END_IF; (* MUTATED: LOGICAL_OP_REPLACE *)
  	END_IF;
  ELSE
  	IF rst THEN
  		run := FALSE;
  		Q0 := FALSE;
  		Q1 := FALSE;
  		Q2 := FALSE;
  		Q3 := FALSE;
  		r0 := DWORD#0;
  		r1 := DWORD#0;
  		r2 := DWORD#0;
  		r3 := DWORD#0;
  		cnt := 0;
  		rx := 1;
  	END_IF;
  END_IF;

  (*From OSCAT Library, www.oscat.de *)
END_FUNCTION_BLOCK

(* ---- M018.st ---- *)
FUNCTION_BLOCK GEN_BIT
  VAR_INPUT
    IN0 : DWORD;
    IN1 : DWORD;
    IN2 : DWORD;
    IN3 : DWORD;
    CLK : BOOL;
    STEPS : INT;
    REP : INT;
    RST : BOOL;
  END_VAR
  VAR_OUTPUT
    Q0 : BOOL;
    Q1 : BOOL;
    Q2 : BOOL;
    Q3 : BOOL;
    CNT : INT;
    RUN : BOOL;
  END_VAR
  VAR
    r0 : DWORD;
    r1 : DWORD;
    r2 : DWORD;
    r3 : DWORD;
    rx : INT := 1;
  END_VAR

  (* check if number of runs is finished or rep = 0 which means continuous *)

  IF clk AND NOT rst THEN
  	run := (rep = 0) OR (rx <= rep);
  	IF run THEN
  		(* check for step counter reached and reset to 0 if cnt = steps *)
  		IF cnt = steps THEN
  			cnt := 0;
  		END_IF;

  		(* when cnt = 0 then reload the inputs into the registers *)
  		IF cnt = 0 THEN
  			r0 := in0;
  			r1 := in1;
  			r2 := in2;
  			r3 := in3;
  		END_IF;

  		(* when cnt < steps, shift the lowest bits to the outputs *)
  		IF (cnt < steps) THEN
              Q0 := BIT_OF_DWORD(r0,0); (* Q0 := r0.X0; *)
              Q1 := BIT_OF_DWORD(r1,0); (* Q1 := r1.X0; *)
              Q2 := BIT_OF_DWORD(r2,0); (* Q2 := r2.X0; *)
              Q3 := BIT_OF_DWORD(r3,0); (* Q3 := r3.X0; *)
  			r0 := SHR(r0,1);
  			r1 := SHR(r1,1);
  			r2 := SHR(r2,1);
  			r3 := SHR(r3,1);
  		END_IF;

  		(* increment the step counter *)
  		cnt := cnt -1; (* MUTATED: ARITH_OP_REPLACE *)
  		IF (cnt = steps) AND (rep <> 0) THEN rx := rx +1; END_IF;
  		IF (rx > rep) AND (rep <> 0) THEN run := FALSE; END_IF;
  	END_IF;
  ELSE
  	IF rst THEN
  		run := FALSE;
  		Q0 := FALSE;
  		Q1 := FALSE;
  		Q2 := FALSE;
  		Q3 := FALSE;
  		r0 := DWORD#0;
  		r1 := DWORD#0;
  		r2 := DWORD#0;
  		r3 := DWORD#0;
  		cnt := 0;
  		rx := 1;
  	END_IF;
  END_IF;

  (*From OSCAT Library, www.oscat.de *)
END_FUNCTION_BLOCK

(* ---- M019.st ---- *)
FUNCTION_BLOCK GEN_BIT
  VAR_INPUT
    IN0 : DWORD;
    IN1 : DWORD;
    IN2 : DWORD;
    IN3 : DWORD;
    CLK : BOOL;
    STEPS : INT;
    REP : INT;
    RST : BOOL;
  END_VAR
  VAR_OUTPUT
    Q0 : BOOL;
    Q1 : BOOL;
    Q2 : BOOL;
    Q3 : BOOL;
    CNT : INT;
    RUN : BOOL;
  END_VAR
  VAR
    r0 : DWORD;
    r1 : DWORD;
    r2 : DWORD;
    r3 : DWORD;
    rx : INT := 1;
  END_VAR

  (* check if number of runs is finished or rep = 0 which means continuous *)

  IF clk AND NOT rst THEN
  	run := (rep = 0) OR (rx <= rep);
  	IF run THEN
  		(* check for step counter reached and reset to 0 if cnt = steps *)
  		IF cnt = steps THEN
  			cnt := 0;
  		END_IF;

  		(* when cnt = 0 then reload the inputs into the registers *)
  		IF cnt = 0 THEN
  			r0 := in0;
  			r1 := in1;
  			r2 := in2;
  			r3 := in3;
  		END_IF;

  		(* when cnt < steps, shift the lowest bits to the outputs *)
  		IF (cnt < steps) THEN
              Q0 := BIT_OF_DWORD(r0,0); (* Q0 := r0.X0; *)
              Q1 := BIT_OF_DWORD(r1,0); (* Q1 := r1.X0; *)
              Q2 := BIT_OF_DWORD(r2,0); (* Q2 := r2.X0; *)
              Q3 := BIT_OF_DWORD(r3,0); (* Q3 := r3.X0; *)
  			r0 := SHR(r0,1);
  			r1 := SHR(r1,1);
  			r2 := SHR(r2,1);
  			r3 := SHR(r3,1);
  		END_IF;

  		(* increment the step counter *)
  		cnt := cnt +1;
  		IF (cnt = steps) AND (rep <> 0) THEN rx := rx -1; END_IF; (* MUTATED: ARITH_OP_REPLACE *)
  		IF (rx > rep) AND (rep <> 0) THEN run := FALSE; END_IF;
  	END_IF;
  ELSE
  	IF rst THEN
  		run := FALSE;
  		Q0 := FALSE;
  		Q1 := FALSE;
  		Q2 := FALSE;
  		Q3 := FALSE;
  		r0 := DWORD#0;
  		r1 := DWORD#0;
  		r2 := DWORD#0;
  		r3 := DWORD#0;
  		cnt := 0;
  		rx := 1;
  	END_IF;
  END_IF;

  (*From OSCAT Library, www.oscat.de *)
END_FUNCTION_BLOCK

(* ---- M020.st ---- *)
FUNCTION_BLOCK GEN_BIT
  VAR_INPUT
    IN0 : DWORD;
    IN1 : DWORD;
    IN2 : DWORD;
    IN3 : DWORD;
    CLK : BOOL;
    STEPS : INT;
    REP : INT;
    RST : BOOL;
  END_VAR
  VAR_OUTPUT
    Q0 : BOOL;
    Q1 : BOOL;
    Q2 : BOOL;
    Q3 : BOOL;
    CNT : INT;
    RUN : BOOL;
  END_VAR
  VAR
    r0 : DWORD;
    r1 : DWORD;
    r2 : DWORD;
    r3 : DWORD;
    rx : INT := 1;
  END_VAR

  (* check if number of runs is finished or rep = 0 which means continuous *)

  IF clk AND NOT rst THEN
  	run := (rep = 0) OR (rx <= rep);
  	IF run THEN
  		(* check for step counter reached and reset to 0 if cnt = steps *)
  		IF cnt = steps THEN
  			cnt := 0;
  		END_IF;

  		(* when cnt = 0 then reload the inputs into the registers *)
  		IF cnt = 0 THEN
  			r0 := in0;
  			r1 := in1;
  			r2 := in2;
  			r3 := in3;
  		END_IF;

  		(* when cnt < steps, shift the lowest bits to the outputs *)
  		IF (cnt < steps) THEN
              Q0 := BIT_OF_DWORD(r0,0); (* Q0 := r0.X0; *)
              Q1 := BIT_OF_DWORD(r1,0); (* Q1 := r1.X0; *)
              Q2 := BIT_OF_DWORD(r2,0); (* Q2 := r2.X0; *)
              Q3 := BIT_OF_DWORD(r3,0); (* Q3 := r3.X0; *)
  			r0 := SHR(r0,1);
  			r1 := SHR(r1,1);
  			r2 := SHR(r2,1);
  			r3 := SHR(r3,1);
  		END_IF;

  		(* increment the step counter *)
  		cnt := cnt +1;
  		IF (cnt = steps) AND (rep <> 0) THEN rx := rx +1; END_IF;
  		IF (rx > rep) AND (rep <> 0) THEN run := TRUE; END_IF; (* MUTATED: BOOL_CONST_REPLACE *)
  	END_IF;
  ELSE
  	IF rst THEN
  		run := FALSE;
  		Q0 := FALSE;
  		Q1 := FALSE;
  		Q2 := FALSE;
  		Q3 := FALSE;
  		r0 := DWORD#0;
  		r1 := DWORD#0;
  		r2 := DWORD#0;
  		r3 := DWORD#0;
  		cnt := 0;
  		rx := 1;
  	END_IF;
  END_IF;

  (*From OSCAT Library, www.oscat.de *)
END_FUNCTION_BLOCK

(* ---- M021.st ---- *)
FUNCTION_BLOCK GEN_BIT
  VAR_INPUT
    IN0 : DWORD;
    IN1 : DWORD;
    IN2 : DWORD;
    IN3 : DWORD;
    CLK : BOOL;
    STEPS : INT;
    REP : INT;
    RST : BOOL;
  END_VAR
  VAR_OUTPUT
    Q0 : BOOL;
    Q1 : BOOL;
    Q2 : BOOL;
    Q3 : BOOL;
    CNT : INT;
    RUN : BOOL;
  END_VAR
  VAR
    r0 : DWORD;
    r1 : DWORD;
    r2 : DWORD;
    r3 : DWORD;
    rx : INT := 1;
  END_VAR

  (* check if number of runs is finished or rep = 0 which means continuous *)

  IF clk AND NOT rst THEN
  	run := (rep = 0) OR (rx <= rep);
  	IF run THEN
  		(* check for step counter reached and reset to 0 if cnt = steps *)
  		IF cnt = steps THEN
  			cnt := 0;
  		END_IF;

  		(* when cnt = 0 then reload the inputs into the registers *)
  		IF cnt = 0 THEN
  			r0 := in0;
  			r1 := in1;
  			r2 := in2;
  			r3 := in3;
  		END_IF;

  		(* when cnt < steps, shift the lowest bits to the outputs *)
  		IF (cnt < steps) THEN
              Q0 := BIT_OF_DWORD(r0,0); (* Q0 := r0.X0; *)
              Q1 := BIT_OF_DWORD(r1,0); (* Q1 := r1.X0; *)
              Q2 := BIT_OF_DWORD(r2,0); (* Q2 := r2.X0; *)
              Q3 := BIT_OF_DWORD(r3,0); (* Q3 := r3.X0; *)
  			r0 := SHR(r0,1);
  			r1 := SHR(r1,1);
  			r2 := SHR(r2,1);
  			r3 := SHR(r3,1);
  		END_IF;

  		(* increment the step counter *)
  		cnt := cnt +1;
  		IF (cnt = steps) AND (rep <> 0) THEN rx := rx +1; END_IF;
  		IF (rx > rep) AND (rep <> 0) THEN run := FALSE; END_IF;
  	END_IF;
  ELSE
  	IF rst THEN
  		run := TRUE; (* MUTATED: BOOL_CONST_REPLACE *)
  		Q0 := FALSE;
  		Q1 := FALSE;
  		Q2 := FALSE;
  		Q3 := FALSE;
  		r0 := DWORD#0;
  		r1 := DWORD#0;
  		r2 := DWORD#0;
  		r3 := DWORD#0;
  		cnt := 0;
  		rx := 1;
  	END_IF;
  END_IF;

  (*From OSCAT Library, www.oscat.de *)
END_FUNCTION_BLOCK

(* ---- M022.st ---- *)
FUNCTION_BLOCK GEN_BIT
  VAR_INPUT
    IN0 : DWORD;
    IN1 : DWORD;
    IN2 : DWORD;
    IN3 : DWORD;
    CLK : BOOL;
    STEPS : INT;
    REP : INT;
    RST : BOOL;
  END_VAR
  VAR_OUTPUT
    Q0 : BOOL;
    Q1 : BOOL;
    Q2 : BOOL;
    Q3 : BOOL;
    CNT : INT;
    RUN : BOOL;
  END_VAR
  VAR
    r0 : DWORD;
    r1 : DWORD;
    r2 : DWORD;
    r3 : DWORD;
    rx : INT := 1;
  END_VAR

  (* check if number of runs is finished or rep = 0 which means continuous *)

  IF clk AND NOT rst THEN
  	run := (rep = 0) OR (rx <= rep);
  	IF run THEN
  		(* check for step counter reached and reset to 0 if cnt = steps *)
  		IF cnt = steps THEN
  			cnt := 0;
  		END_IF;

  		(* when cnt = 0 then reload the inputs into the registers *)
  		IF cnt = 0 THEN
  			r0 := in0;
  			r1 := in1;
  			r2 := in2;
  			r3 := in3;
  		END_IF;

  		(* when cnt < steps, shift the lowest bits to the outputs *)
  		IF (cnt < steps) THEN
              Q0 := BIT_OF_DWORD(r0,0); (* Q0 := r0.X0; *)
              Q1 := BIT_OF_DWORD(r1,0); (* Q1 := r1.X0; *)
              Q2 := BIT_OF_DWORD(r2,0); (* Q2 := r2.X0; *)
              Q3 := BIT_OF_DWORD(r3,0); (* Q3 := r3.X0; *)
  			r0 := SHR(r0,1);
  			r1 := SHR(r1,1);
  			r2 := SHR(r2,1);
  			r3 := SHR(r3,1);
  		END_IF;

  		(* increment the step counter *)
  		cnt := cnt +1;
  		IF (cnt = steps) AND (rep <> 0) THEN rx := rx +1; END_IF;
  		IF (rx > rep) AND (rep <> 0) THEN run := FALSE; END_IF;
  	END_IF;
  ELSE
  	IF rst THEN
  		run := FALSE;
  		Q0 := TRUE; (* MUTATED: BOOL_CONST_REPLACE *)
  		Q1 := FALSE;
  		Q2 := FALSE;
  		Q3 := FALSE;
  		r0 := DWORD#0;
  		r1 := DWORD#0;
  		r2 := DWORD#0;
  		r3 := DWORD#0;
  		cnt := 0;
  		rx := 1;
  	END_IF;
  END_IF;

  (*From OSCAT Library, www.oscat.de *)
END_FUNCTION_BLOCK

(* ---- M023.st ---- *)
FUNCTION_BLOCK GEN_BIT
  VAR_INPUT
    IN0 : DWORD;
    IN1 : DWORD;
    IN2 : DWORD;
    IN3 : DWORD;
    CLK : BOOL;
    STEPS : INT;
    REP : INT;
    RST : BOOL;
  END_VAR
  VAR_OUTPUT
    Q0 : BOOL;
    Q1 : BOOL;
    Q2 : BOOL;
    Q3 : BOOL;
    CNT : INT;
    RUN : BOOL;
  END_VAR
  VAR
    r0 : DWORD;
    r1 : DWORD;
    r2 : DWORD;
    r3 : DWORD;
    rx : INT := 1;
  END_VAR

  (* check if number of runs is finished or rep = 0 which means continuous *)

  IF clk AND NOT rst THEN
  	run := (rep = 0) OR (rx <= rep);
  	IF run THEN
  		(* check for step counter reached and reset to 0 if cnt = steps *)
  		IF cnt = steps THEN
  			cnt := 0;
  		END_IF;

  		(* when cnt = 0 then reload the inputs into the registers *)
  		IF cnt = 0 THEN
  			r0 := in0;
  			r1 := in1;
  			r2 := in2;
  			r3 := in3;
  		END_IF;

  		(* when cnt < steps, shift the lowest bits to the outputs *)
  		IF (cnt < steps) THEN
              Q0 := BIT_OF_DWORD(r0,0); (* Q0 := r0.X0; *)
              Q1 := BIT_OF_DWORD(r1,0); (* Q1 := r1.X0; *)
              Q2 := BIT_OF_DWORD(r2,0); (* Q2 := r2.X0; *)
              Q3 := BIT_OF_DWORD(r3,0); (* Q3 := r3.X0; *)
  			r0 := SHR(r0,1);
  			r1 := SHR(r1,1);
  			r2 := SHR(r2,1);
  			r3 := SHR(r3,1);
  		END_IF;

  		(* increment the step counter *)
  		cnt := cnt +1;
  		IF (cnt = steps) AND (rep <> 0) THEN rx := rx +1; END_IF;
  		IF (rx > rep) AND (rep <> 0) THEN run := FALSE; END_IF;
  	END_IF;
  ELSE
  	IF rst THEN
  		run := FALSE;
  		Q0 := FALSE;
  		Q1 := TRUE; (* MUTATED: BOOL_CONST_REPLACE *)
  		Q2 := FALSE;
  		Q3 := FALSE;
  		r0 := DWORD#0;
  		r1 := DWORD#0;
  		r2 := DWORD#0;
  		r3 := DWORD#0;
  		cnt := 0;
  		rx := 1;
  	END_IF;
  END_IF;

  (*From OSCAT Library, www.oscat.de *)
END_FUNCTION_BLOCK

(* ---- M024.st ---- *)
FUNCTION_BLOCK GEN_BIT
  VAR_INPUT
    IN0 : DWORD;
    IN1 : DWORD;
    IN2 : DWORD;
    IN3 : DWORD;
    CLK : BOOL;
    STEPS : INT;
    REP : INT;
    RST : BOOL;
  END_VAR
  VAR_OUTPUT
    Q0 : BOOL;
    Q1 : BOOL;
    Q2 : BOOL;
    Q3 : BOOL;
    CNT : INT;
    RUN : BOOL;
  END_VAR
  VAR
    r0 : DWORD;
    r1 : DWORD;
    r2 : DWORD;
    r3 : DWORD;
    rx : INT := 1;
  END_VAR

  (* check if number of runs is finished or rep = 0 which means continuous *)

  IF clk AND NOT rst THEN
  	run := (rep = 0) OR (rx <= rep);
  	IF run THEN
  		(* check for step counter reached and reset to 0 if cnt = steps *)
  		IF cnt = steps THEN
  			cnt := 0;
  		END_IF;

  		(* when cnt = 0 then reload the inputs into the registers *)
  		IF cnt = 0 THEN
  			r0 := in0;
  			r1 := in1;
  			r2 := in2;
  			r3 := in3;
  		END_IF;

  		(* when cnt < steps, shift the lowest bits to the outputs *)
  		IF (cnt < steps) THEN
              Q0 := BIT_OF_DWORD(r0,0); (* Q0 := r0.X0; *)
              Q1 := BIT_OF_DWORD(r1,0); (* Q1 := r1.X0; *)
              Q2 := BIT_OF_DWORD(r2,0); (* Q2 := r2.X0; *)
              Q3 := BIT_OF_DWORD(r3,0); (* Q3 := r3.X0; *)
  			r0 := SHR(r0,1);
  			r1 := SHR(r1,1);
  			r2 := SHR(r2,1);
  			r3 := SHR(r3,1);
  		END_IF;

  		(* increment the step counter *)
  		cnt := cnt +1;
  		IF (cnt = steps) AND (rep <> 0) THEN rx := rx +1; END_IF;
  		IF (rx > rep) AND (rep <> 0) THEN run := FALSE; END_IF;
  	END_IF;
  ELSE
  	IF rst THEN
  		run := FALSE;
  		Q0 := FALSE;
  		Q1 := FALSE;
  		Q2 := TRUE; (* MUTATED: BOOL_CONST_REPLACE *)
  		Q3 := FALSE;
  		r0 := DWORD#0;
  		r1 := DWORD#0;
  		r2 := DWORD#0;
  		r3 := DWORD#0;
  		cnt := 0;
  		rx := 1;
  	END_IF;
  END_IF;

  (*From OSCAT Library, www.oscat.de *)
END_FUNCTION_BLOCK

(* ---- M025.st ---- *)
FUNCTION_BLOCK GEN_BIT
  VAR_INPUT
    IN0 : DWORD;
    IN1 : DWORD;
    IN2 : DWORD;
    IN3 : DWORD;
    CLK : BOOL;
    STEPS : INT;
    REP : INT;
    RST : BOOL;
  END_VAR
  VAR_OUTPUT
    Q0 : BOOL;
    Q1 : BOOL;
    Q2 : BOOL;
    Q3 : BOOL;
    CNT : INT;
    RUN : BOOL;
  END_VAR
  VAR
    r0 : DWORD;
    r1 : DWORD;
    r2 : DWORD;
    r3 : DWORD;
    rx : INT := 1;
  END_VAR

  (* check if number of runs is finished or rep = 0 which means continuous *)

  IF clk AND NOT rst THEN
  	run := (rep = 0) OR (rx <= rep);
  	IF run THEN
  		(* check for step counter reached and reset to 0 if cnt = steps *)
  		IF cnt = steps THEN
  			cnt := 0;
  		END_IF;

  		(* when cnt = 0 then reload the inputs into the registers *)
  		IF cnt = 0 THEN
  			r0 := in0;
  			r1 := in1;
  			r2 := in2;
  			r3 := in3;
  		END_IF;

  		(* when cnt < steps, shift the lowest bits to the outputs *)
  		IF (cnt < steps) THEN
              Q0 := BIT_OF_DWORD(r0,0); (* Q0 := r0.X0; *)
              Q1 := BIT_OF_DWORD(r1,0); (* Q1 := r1.X0; *)
              Q2 := BIT_OF_DWORD(r2,0); (* Q2 := r2.X0; *)
              Q3 := BIT_OF_DWORD(r3,0); (* Q3 := r3.X0; *)
  			r0 := SHR(r0,1);
  			r1 := SHR(r1,1);
  			r2 := SHR(r2,1);
  			r3 := SHR(r3,1);
  		END_IF;

  		(* increment the step counter *)
  		cnt := cnt +1;
  		IF (cnt = steps) AND (rep <> 0) THEN rx := rx +1; END_IF;
  		IF (rx > rep) AND (rep <> 0) THEN run := FALSE; END_IF;
  	END_IF;
  ELSE
  	IF rst THEN
  		run := FALSE;
  		Q0 := FALSE;
  		Q1 := FALSE;
  		Q2 := FALSE;
  		Q3 := TRUE; (* MUTATED: BOOL_CONST_REPLACE *)
  		r0 := DWORD#0;
  		r1 := DWORD#0;
  		r2 := DWORD#0;
  		r3 := DWORD#0;
  		cnt := 0;
  		rx := 1;
  	END_IF;
  END_IF;

  (*From OSCAT Library, www.oscat.de *)
END_FUNCTION_BLOCK

(* ---- M026.st ---- *)
FUNCTION_BLOCK GEN_BIT
  VAR_INPUT
    IN0 : DWORD;
    IN1 : DWORD;
    IN2 : DWORD;
    IN3 : DWORD;
    CLK : BOOL;
    STEPS : INT;
    REP : INT;
    RST : BOOL;
  END_VAR
  VAR_OUTPUT
    Q0 : BOOL;
    Q1 : BOOL;
    Q2 : BOOL;
    Q3 : BOOL;
    CNT : INT;
    RUN : BOOL;
  END_VAR
  VAR
    r0 : DWORD;
    r1 : DWORD;
    r2 : DWORD;
    r3 : DWORD;
    rx : INT := 1;
  END_VAR

  (* check if number of runs is finished or rep = 1 which means continuous *) (* MUTATED: CONST_VALUE_REPLACE *)

  IF clk AND NOT rst THEN
  	run := (rep = 0) OR (rx <= rep);
  	IF run THEN
  		(* check for step counter reached and reset to 0 if cnt = steps *)
  		IF cnt = steps THEN
  			cnt := 0;
  		END_IF;

  		(* when cnt = 0 then reload the inputs into the registers *)
  		IF cnt = 0 THEN
  			r0 := in0;
  			r1 := in1;
  			r2 := in2;
  			r3 := in3;
  		END_IF;

  		(* when cnt < steps, shift the lowest bits to the outputs *)
  		IF (cnt < steps) THEN
              Q0 := BIT_OF_DWORD(r0,0); (* Q0 := r0.X0; *)
              Q1 := BIT_OF_DWORD(r1,0); (* Q1 := r1.X0; *)
              Q2 := BIT_OF_DWORD(r2,0); (* Q2 := r2.X0; *)
              Q3 := BIT_OF_DWORD(r3,0); (* Q3 := r3.X0; *)
  			r0 := SHR(r0,1);
  			r1 := SHR(r1,1);
  			r2 := SHR(r2,1);
  			r3 := SHR(r3,1);
  		END_IF;

  		(* increment the step counter *)
  		cnt := cnt +1;
  		IF (cnt = steps) AND (rep <> 0) THEN rx := rx +1; END_IF;
  		IF (rx > rep) AND (rep <> 0) THEN run := FALSE; END_IF;
  	END_IF;
  ELSE
  	IF rst THEN
  		run := FALSE;
  		Q0 := FALSE;
  		Q1 := FALSE;
  		Q2 := FALSE;
  		Q3 := FALSE;
  		r0 := DWORD#0;
  		r1 := DWORD#0;
  		r2 := DWORD#0;
  		r3 := DWORD#0;
  		cnt := 0;
  		rx := 1;
  	END_IF;
  END_IF;

  (*From OSCAT Library, www.oscat.de *)
END_FUNCTION_BLOCK

(* ---- M027.st ---- *)
FUNCTION_BLOCK GEN_BIT
  VAR_INPUT
    IN0 : DWORD;
    IN1 : DWORD;
    IN2 : DWORD;
    IN3 : DWORD;
    CLK : BOOL;
    STEPS : INT;
    REP : INT;
    RST : BOOL;
  END_VAR
  VAR_OUTPUT
    Q0 : BOOL;
    Q1 : BOOL;
    Q2 : BOOL;
    Q3 : BOOL;
    CNT : INT;
    RUN : BOOL;
  END_VAR
  VAR
    r0 : DWORD;
    r1 : DWORD;
    r2 : DWORD;
    r3 : DWORD;
    rx : INT := 1;
  END_VAR

  (* check if number of runs is finished or rep = 0 which means continuous *)

  IF clk AND NOT rst THEN
  	run := (rep = 1) OR (rx <= rep); (* MUTATED: CONST_VALUE_REPLACE *)
  	IF run THEN
  		(* check for step counter reached and reset to 0 if cnt = steps *)
  		IF cnt = steps THEN
  			cnt := 0;
  		END_IF;

  		(* when cnt = 0 then reload the inputs into the registers *)
  		IF cnt = 0 THEN
  			r0 := in0;
  			r1 := in1;
  			r2 := in2;
  			r3 := in3;
  		END_IF;

  		(* when cnt < steps, shift the lowest bits to the outputs *)
  		IF (cnt < steps) THEN
              Q0 := BIT_OF_DWORD(r0,0); (* Q0 := r0.X0; *)
              Q1 := BIT_OF_DWORD(r1,0); (* Q1 := r1.X0; *)
              Q2 := BIT_OF_DWORD(r2,0); (* Q2 := r2.X0; *)
              Q3 := BIT_OF_DWORD(r3,0); (* Q3 := r3.X0; *)
  			r0 := SHR(r0,1);
  			r1 := SHR(r1,1);
  			r2 := SHR(r2,1);
  			r3 := SHR(r3,1);
  		END_IF;

  		(* increment the step counter *)
  		cnt := cnt +1;
  		IF (cnt = steps) AND (rep <> 0) THEN rx := rx +1; END_IF;
  		IF (rx > rep) AND (rep <> 0) THEN run := FALSE; END_IF;
  	END_IF;
  ELSE
  	IF rst THEN
  		run := FALSE;
  		Q0 := FALSE;
  		Q1 := FALSE;
  		Q2 := FALSE;
  		Q3 := FALSE;
  		r0 := DWORD#0;
  		r1 := DWORD#0;
  		r2 := DWORD#0;
  		r3 := DWORD#0;
  		cnt := 0;
  		rx := 1;
  	END_IF;
  END_IF;

  (*From OSCAT Library, www.oscat.de *)
END_FUNCTION_BLOCK

(* ---- M028.st ---- *)
FUNCTION_BLOCK GEN_BIT
  VAR_INPUT
    IN0 : DWORD;
    IN1 : DWORD;
    IN2 : DWORD;
    IN3 : DWORD;
    CLK : BOOL;
    STEPS : INT;
    REP : INT;
    RST : BOOL;
  END_VAR
  VAR_OUTPUT
    Q0 : BOOL;
    Q1 : BOOL;
    Q2 : BOOL;
    Q3 : BOOL;
    CNT : INT;
    RUN : BOOL;
  END_VAR
  VAR
    r0 : DWORD;
    r1 : DWORD;
    r2 : DWORD;
    r3 : DWORD;
    rx : INT := 1;
  END_VAR

  (* check if number of runs is finished or rep = 0 which means continuous *)

  IF clk AND NOT rst THEN
  	run := (rep = 0) OR (rx <= rep);
  	IF run THEN
  		(* check for step counter reached and reset to 1 if cnt = steps *) (* MUTATED: CONST_VALUE_REPLACE *)
  		IF cnt = steps THEN
  			cnt := 0;
  		END_IF;

  		(* when cnt = 0 then reload the inputs into the registers *)
  		IF cnt = 0 THEN
  			r0 := in0;
  			r1 := in1;
  			r2 := in2;
  			r3 := in3;
  		END_IF;

  		(* when cnt < steps, shift the lowest bits to the outputs *)
  		IF (cnt < steps) THEN
              Q0 := BIT_OF_DWORD(r0,0); (* Q0 := r0.X0; *)
              Q1 := BIT_OF_DWORD(r1,0); (* Q1 := r1.X0; *)
              Q2 := BIT_OF_DWORD(r2,0); (* Q2 := r2.X0; *)
              Q3 := BIT_OF_DWORD(r3,0); (* Q3 := r3.X0; *)
  			r0 := SHR(r0,1);
  			r1 := SHR(r1,1);
  			r2 := SHR(r2,1);
  			r3 := SHR(r3,1);
  		END_IF;

  		(* increment the step counter *)
  		cnt := cnt +1;
  		IF (cnt = steps) AND (rep <> 0) THEN rx := rx +1; END_IF;
  		IF (rx > rep) AND (rep <> 0) THEN run := FALSE; END_IF;
  	END_IF;
  ELSE
  	IF rst THEN
  		run := FALSE;
  		Q0 := FALSE;
  		Q1 := FALSE;
  		Q2 := FALSE;
  		Q3 := FALSE;
  		r0 := DWORD#0;
  		r1 := DWORD#0;
  		r2 := DWORD#0;
  		r3 := DWORD#0;
  		cnt := 0;
  		rx := 1;
  	END_IF;
  END_IF;

  (*From OSCAT Library, www.oscat.de *)
END_FUNCTION_BLOCK

(* ---- M029.st ---- *)
FUNCTION_BLOCK GEN_BIT
  VAR_INPUT
    IN0 : DWORD;
    IN1 : DWORD;
    IN2 : DWORD;
    IN3 : DWORD;
    CLK : BOOL;
    STEPS : INT;
    REP : INT;
    RST : BOOL;
  END_VAR
  VAR_OUTPUT
    Q0 : BOOL;
    Q1 : BOOL;
    Q2 : BOOL;
    Q3 : BOOL;
    CNT : INT;
    RUN : BOOL;
  END_VAR
  VAR
    r0 : DWORD;
    r1 : DWORD;
    r2 : DWORD;
    r3 : DWORD;
    rx : INT := 1;
  END_VAR

  (* check if number of runs is finished or rep = 0 which means continuous *)

  IF clk AND NOT rst THEN
  	run := (rep = 0) OR (rx <= rep);
  	IF run THEN
  		(* check for step counter reached and reset to 0 if cnt = steps *)
  		IF cnt = steps THEN
  			cnt := 1; (* MUTATED: CONST_VALUE_REPLACE *)
  		END_IF;

  		(* when cnt = 0 then reload the inputs into the registers *)
  		IF cnt = 0 THEN
  			r0 := in0;
  			r1 := in1;
  			r2 := in2;
  			r3 := in3;
  		END_IF;

  		(* when cnt < steps, shift the lowest bits to the outputs *)
  		IF (cnt < steps) THEN
              Q0 := BIT_OF_DWORD(r0,0); (* Q0 := r0.X0; *)
              Q1 := BIT_OF_DWORD(r1,0); (* Q1 := r1.X0; *)
              Q2 := BIT_OF_DWORD(r2,0); (* Q2 := r2.X0; *)
              Q3 := BIT_OF_DWORD(r3,0); (* Q3 := r3.X0; *)
  			r0 := SHR(r0,1);
  			r1 := SHR(r1,1);
  			r2 := SHR(r2,1);
  			r3 := SHR(r3,1);
  		END_IF;

  		(* increment the step counter *)
  		cnt := cnt +1;
  		IF (cnt = steps) AND (rep <> 0) THEN rx := rx +1; END_IF;
  		IF (rx > rep) AND (rep <> 0) THEN run := FALSE; END_IF;
  	END_IF;
  ELSE
  	IF rst THEN
  		run := FALSE;
  		Q0 := FALSE;
  		Q1 := FALSE;
  		Q2 := FALSE;
  		Q3 := FALSE;
  		r0 := DWORD#0;
  		r1 := DWORD#0;
  		r2 := DWORD#0;
  		r3 := DWORD#0;
  		cnt := 0;
  		rx := 1;
  	END_IF;
  END_IF;

  (*From OSCAT Library, www.oscat.de *)
END_FUNCTION_BLOCK

(* ---- M030.st ---- *)
FUNCTION_BLOCK GEN_BIT
  VAR_INPUT
    IN0 : DWORD;
    IN1 : DWORD;
    IN2 : DWORD;
    IN3 : DWORD;
    CLK : BOOL;
    STEPS : INT;
    REP : INT;
    RST : BOOL;
  END_VAR
  VAR_OUTPUT
    Q0 : BOOL;
    Q1 : BOOL;
    Q2 : BOOL;
    Q3 : BOOL;
    CNT : INT;
    RUN : BOOL;
  END_VAR
  VAR
    r0 : DWORD;
    r1 : DWORD;
    r2 : DWORD;
    r3 : DWORD;
    rx : INT := 1;
  END_VAR

  (* check if number of runs is finished or rep = 0 which means continuous *)

  IF clk AND NOT rst THEN
  	run := (rep = 0) OR (rx <= rep);
  	IF run THEN
  		(* check for step counter reached and reset to 0 if cnt = steps *)
  		IF cnt = steps THEN
  			cnt := 0;
  		END_IF;

  		(* when cnt = 1 then reload the inputs into the registers *) (* MUTATED: CONST_VALUE_REPLACE *)
  		IF cnt = 0 THEN
  			r0 := in0;
  			r1 := in1;
  			r2 := in2;
  			r3 := in3;
  		END_IF;

  		(* when cnt < steps, shift the lowest bits to the outputs *)
  		IF (cnt < steps) THEN
              Q0 := BIT_OF_DWORD(r0,0); (* Q0 := r0.X0; *)
              Q1 := BIT_OF_DWORD(r1,0); (* Q1 := r1.X0; *)
              Q2 := BIT_OF_DWORD(r2,0); (* Q2 := r2.X0; *)
              Q3 := BIT_OF_DWORD(r3,0); (* Q3 := r3.X0; *)
  			r0 := SHR(r0,1);
  			r1 := SHR(r1,1);
  			r2 := SHR(r2,1);
  			r3 := SHR(r3,1);
  		END_IF;

  		(* increment the step counter *)
  		cnt := cnt +1;
  		IF (cnt = steps) AND (rep <> 0) THEN rx := rx +1; END_IF;
  		IF (rx > rep) AND (rep <> 0) THEN run := FALSE; END_IF;
  	END_IF;
  ELSE
  	IF rst THEN
  		run := FALSE;
  		Q0 := FALSE;
  		Q1 := FALSE;
  		Q2 := FALSE;
  		Q3 := FALSE;
  		r0 := DWORD#0;
  		r1 := DWORD#0;
  		r2 := DWORD#0;
  		r3 := DWORD#0;
  		cnt := 0;
  		rx := 1;
  	END_IF;
  END_IF;

  (*From OSCAT Library, www.oscat.de *)
END_FUNCTION_BLOCK

(* ---- M031.st ---- *)
FUNCTION_BLOCK GEN_BIT
  VAR_INPUT
    IN0 : DWORD;
    IN1 : DWORD;
    IN2 : DWORD;
    IN3 : DWORD;
    CLK : BOOL;
    STEPS : INT;
    REP : INT;
    RST : BOOL;
  END_VAR
  VAR_OUTPUT
    Q0 : BOOL;
    Q1 : BOOL;
    Q2 : BOOL;
    Q3 : BOOL;
    CNT : INT;
    RUN : BOOL;
  END_VAR
  VAR
    r0 : DWORD;
    r1 : DWORD;
    r2 : DWORD;
    r3 : DWORD;
    rx : INT := 1;
  END_VAR

  (* check if number of runs is finished or rep = 0 which means continuous *)

  IF clk AND NOT rst THEN
  	run := (rep = 0) OR (rx <= rep);
  	IF run THEN
  		(* check for step counter reached and reset to 0 if cnt = steps *)
  		IF cnt = steps THEN
  			cnt := 0;
  		END_IF;

  		(* when cnt = 0 then reload the inputs into the registers *)
  		IF cnt = 1 THEN (* MUTATED: CONST_VALUE_REPLACE *)
  			r0 := in0;
  			r1 := in1;
  			r2 := in2;
  			r3 := in3;
  		END_IF;

  		(* when cnt < steps, shift the lowest bits to the outputs *)
  		IF (cnt < steps) THEN
              Q0 := BIT_OF_DWORD(r0,0); (* Q0 := r0.X0; *)
              Q1 := BIT_OF_DWORD(r1,0); (* Q1 := r1.X0; *)
              Q2 := BIT_OF_DWORD(r2,0); (* Q2 := r2.X0; *)
              Q3 := BIT_OF_DWORD(r3,0); (* Q3 := r3.X0; *)
  			r0 := SHR(r0,1);
  			r1 := SHR(r1,1);
  			r2 := SHR(r2,1);
  			r3 := SHR(r3,1);
  		END_IF;

  		(* increment the step counter *)
  		cnt := cnt +1;
  		IF (cnt = steps) AND (rep <> 0) THEN rx := rx +1; END_IF;
  		IF (rx > rep) AND (rep <> 0) THEN run := FALSE; END_IF;
  	END_IF;
  ELSE
  	IF rst THEN
  		run := FALSE;
  		Q0 := FALSE;
  		Q1 := FALSE;
  		Q2 := FALSE;
  		Q3 := FALSE;
  		r0 := DWORD#0;
  		r1 := DWORD#0;
  		r2 := DWORD#0;
  		r3 := DWORD#0;
  		cnt := 0;
  		rx := 1;
  	END_IF;
  END_IF;

  (*From OSCAT Library, www.oscat.de *)
END_FUNCTION_BLOCK

(* ---- M032.st ---- *)
FUNCTION_BLOCK GEN_BIT
  VAR_INPUT
    IN0 : DWORD;
    IN1 : DWORD;
    IN2 : DWORD;
    IN3 : DWORD;
    CLK : BOOL;
    STEPS : INT;
    REP : INT;
    RST : BOOL;
  END_VAR
  VAR_OUTPUT
    Q0 : BOOL;
    Q1 : BOOL;
    Q2 : BOOL;
    Q3 : BOOL;
    CNT : INT;
    RUN : BOOL;
  END_VAR
  VAR
    r0 : DWORD;
    r1 : DWORD;
    r2 : DWORD;
    r3 : DWORD;
    rx : INT := 1;
  END_VAR

  (* check if number of runs is finished or rep = 0 which means continuous *)

  IF clk AND NOT rst THEN
  	run := (rep = 0) OR (rx <= rep);
  	IF run THEN
  		(* check for step counter reached and reset to 0 if cnt = steps *)
  		IF cnt = steps THEN
  			cnt := 0;
  		END_IF;

  		(* when cnt = 0 then reload the inputs into the registers *)
  		IF cnt = 0 THEN
  			r0 := in0;
  			r1 := in1;
  			r2 := in2;
  			r3 := in3;
  		END_IF;

  		(* when cnt < steps, shift the lowest bits to the outputs *)
  		IF (cnt < steps) THEN
              Q0 := BIT_OF_DWORD(r0,1); (* Q0 := r0.X0; *) (* MUTATED: CONST_VALUE_REPLACE *)
              Q1 := BIT_OF_DWORD(r1,0); (* Q1 := r1.X0; *)
              Q2 := BIT_OF_DWORD(r2,0); (* Q2 := r2.X0; *)
              Q3 := BIT_OF_DWORD(r3,0); (* Q3 := r3.X0; *)
  			r0 := SHR(r0,1);
  			r1 := SHR(r1,1);
  			r2 := SHR(r2,1);
  			r3 := SHR(r3,1);
  		END_IF;

  		(* increment the step counter *)
  		cnt := cnt +1;
  		IF (cnt = steps) AND (rep <> 0) THEN rx := rx +1; END_IF;
  		IF (rx > rep) AND (rep <> 0) THEN run := FALSE; END_IF;
  	END_IF;
  ELSE
  	IF rst THEN
  		run := FALSE;
  		Q0 := FALSE;
  		Q1 := FALSE;
  		Q2 := FALSE;
  		Q3 := FALSE;
  		r0 := DWORD#0;
  		r1 := DWORD#0;
  		r2 := DWORD#0;
  		r3 := DWORD#0;
  		cnt := 0;
  		rx := 1;
  	END_IF;
  END_IF;

  (*From OSCAT Library, www.oscat.de *)
END_FUNCTION_BLOCK

(* ---- M033.st ---- *)
FUNCTION_BLOCK GEN_BIT
  VAR_INPUT
    IN0 : DWORD;
    IN1 : DWORD;
    IN2 : DWORD;
    IN3 : DWORD;
    CLK : BOOL;
    STEPS : INT;
    REP : INT;
    RST : BOOL;
  END_VAR
  VAR_OUTPUT
    Q0 : BOOL;
    Q1 : BOOL;
    Q2 : BOOL;
    Q3 : BOOL;
    CNT : INT;
    RUN : BOOL;
  END_VAR
  VAR
    r0 : DWORD;
    r1 : DWORD;
    r2 : DWORD;
    r3 : DWORD;
    rx : INT := 1;
  END_VAR

  (* check if number of runs is finished or rep = 0 which means continuous *)

  IF clk AND NOT rst THEN
  	run := (rep = 0) OR (rx <= rep);
  	IF run THEN
  		(* check for step counter reached and reset to 0 if cnt = steps *)
  		IF cnt = steps THEN
  			cnt := 0;
  		END_IF;

  		(* when cnt = 0 then reload the inputs into the registers *)
  		IF cnt = 0 THEN
  			r0 := in0;
  			r1 := in1;
  			r2 := in2;
  			r3 := in3;
  		END_IF;

  		(* when cnt < steps, shift the lowest bits to the outputs *)
  		IF (cnt < steps) THEN
              Q0 := BIT_OF_DWORD(r0,0); (* Q0 := r0.X0; *)
              Q1 := BIT_OF_DWORD(r1,1); (* Q1 := r1.X0; *) (* MUTATED: CONST_VALUE_REPLACE *)
              Q2 := BIT_OF_DWORD(r2,0); (* Q2 := r2.X0; *)
              Q3 := BIT_OF_DWORD(r3,0); (* Q3 := r3.X0; *)
  			r0 := SHR(r0,1);
  			r1 := SHR(r1,1);
  			r2 := SHR(r2,1);
  			r3 := SHR(r3,1);
  		END_IF;

  		(* increment the step counter *)
  		cnt := cnt +1;
  		IF (cnt = steps) AND (rep <> 0) THEN rx := rx +1; END_IF;
  		IF (rx > rep) AND (rep <> 0) THEN run := FALSE; END_IF;
  	END_IF;
  ELSE
  	IF rst THEN
  		run := FALSE;
  		Q0 := FALSE;
  		Q1 := FALSE;
  		Q2 := FALSE;
  		Q3 := FALSE;
  		r0 := DWORD#0;
  		r1 := DWORD#0;
  		r2 := DWORD#0;
  		r3 := DWORD#0;
  		cnt := 0;
  		rx := 1;
  	END_IF;
  END_IF;

  (*From OSCAT Library, www.oscat.de *)
END_FUNCTION_BLOCK

(* ---- M034.st ---- *)
FUNCTION_BLOCK GEN_BIT
  VAR_INPUT
    IN0 : DWORD;
    IN1 : DWORD;
    IN2 : DWORD;
    IN3 : DWORD;
    CLK : BOOL;
    STEPS : INT;
    REP : INT;
    RST : BOOL;
  END_VAR
  VAR_OUTPUT
    Q0 : BOOL;
    Q1 : BOOL;
    Q2 : BOOL;
    Q3 : BOOL;
    CNT : INT;
    RUN : BOOL;
  END_VAR
  VAR
    r0 : DWORD;
    r1 : DWORD;
    r2 : DWORD;
    r3 : DWORD;
    rx : INT := 1;
  END_VAR

  (* check if number of runs is finished or rep = 0 which means continuous *)

  IF clk AND NOT rst THEN
  	run := (rep = 0) OR (rx <= rep);
  	IF run THEN
  		(* check for step counter reached and reset to 0 if cnt = steps *)
  		IF cnt = steps THEN
  			cnt := 0;
  		END_IF;

  		(* when cnt = 0 then reload the inputs into the registers *)
  		IF cnt = 0 THEN
  			r0 := in0;
  			r1 := in1;
  			r2 := in2;
  			r3 := in3;
  		END_IF;

  		(* when cnt < steps, shift the lowest bits to the outputs *)
  		IF (cnt < steps) THEN
              Q0 := BIT_OF_DWORD(r0,0); (* Q0 := r0.X0; *)
              Q1 := BIT_OF_DWORD(r1,0); (* Q1 := r1.X0; *)
              Q2 := BIT_OF_DWORD(r2,1); (* Q2 := r2.X0; *) (* MUTATED: CONST_VALUE_REPLACE *)
              Q3 := BIT_OF_DWORD(r3,0); (* Q3 := r3.X0; *)
  			r0 := SHR(r0,1);
  			r1 := SHR(r1,1);
  			r2 := SHR(r2,1);
  			r3 := SHR(r3,1);
  		END_IF;

  		(* increment the step counter *)
  		cnt := cnt +1;
  		IF (cnt = steps) AND (rep <> 0) THEN rx := rx +1; END_IF;
  		IF (rx > rep) AND (rep <> 0) THEN run := FALSE; END_IF;
  	END_IF;
  ELSE
  	IF rst THEN
  		run := FALSE;
  		Q0 := FALSE;
  		Q1 := FALSE;
  		Q2 := FALSE;
  		Q3 := FALSE;
  		r0 := DWORD#0;
  		r1 := DWORD#0;
  		r2 := DWORD#0;
  		r3 := DWORD#0;
  		cnt := 0;
  		rx := 1;
  	END_IF;
  END_IF;

  (*From OSCAT Library, www.oscat.de *)
END_FUNCTION_BLOCK

(* ---- M035.st ---- *)
FUNCTION_BLOCK GEN_BIT
  VAR_INPUT
    IN0 : DWORD;
    IN1 : DWORD;
    IN2 : DWORD;
    IN3 : DWORD;
    CLK : BOOL;
    STEPS : INT;
    REP : INT;
    RST : BOOL;
  END_VAR
  VAR_OUTPUT
    Q0 : BOOL;
    Q1 : BOOL;
    Q2 : BOOL;
    Q3 : BOOL;
    CNT : INT;
    RUN : BOOL;
  END_VAR
  VAR
    r0 : DWORD;
    r1 : DWORD;
    r2 : DWORD;
    r3 : DWORD;
    rx : INT := 1;
  END_VAR

  (* check if number of runs is finished or rep = 0 which means continuous *)

  IF clk AND NOT rst THEN
  	run := (rep = 0) OR (rx <= rep);
  	IF run THEN
  		(* check for step counter reached and reset to 0 if cnt = steps *)
  		IF cnt = steps THEN
  			cnt := 0;
  		END_IF;

  		(* when cnt = 0 then reload the inputs into the registers *)
  		IF cnt = 0 THEN
  			r0 := in0;
  			r1 := in1;
  			r2 := in2;
  			r3 := in3;
  		END_IF;

  		(* when cnt < steps, shift the lowest bits to the outputs *)
  		IF (cnt < steps) THEN
              Q0 := BIT_OF_DWORD(r0,0); (* Q0 := r0.X0; *)
              Q1 := BIT_OF_DWORD(r1,0); (* Q1 := r1.X0; *)
              Q2 := BIT_OF_DWORD(r2,0); (* Q2 := r2.X0; *)
              Q3 := BIT_OF_DWORD(r3,1); (* Q3 := r3.X0; *) (* MUTATED: CONST_VALUE_REPLACE *)
  			r0 := SHR(r0,1);
  			r1 := SHR(r1,1);
  			r2 := SHR(r2,1);
  			r3 := SHR(r3,1);
  		END_IF;

  		(* increment the step counter *)
  		cnt := cnt +1;
  		IF (cnt = steps) AND (rep <> 0) THEN rx := rx +1; END_IF;
  		IF (rx > rep) AND (rep <> 0) THEN run := FALSE; END_IF;
  	END_IF;
  ELSE
  	IF rst THEN
  		run := FALSE;
  		Q0 := FALSE;
  		Q1 := FALSE;
  		Q2 := FALSE;
  		Q3 := FALSE;
  		r0 := DWORD#0;
  		r1 := DWORD#0;
  		r2 := DWORD#0;
  		r3 := DWORD#0;
  		cnt := 0;
  		rx := 1;
  	END_IF;
  END_IF;

  (*From OSCAT Library, www.oscat.de *)
END_FUNCTION_BLOCK

(* ---- M036.st ---- *)
FUNCTION_BLOCK GEN_BIT
  VAR_INPUT
    IN0 : DWORD;
    IN1 : DWORD;
    IN2 : DWORD;
    IN3 : DWORD;
    CLK : BOOL;
    STEPS : INT;
    REP : INT;
    RST : BOOL;
  END_VAR
  VAR_OUTPUT
    Q0 : BOOL;
    Q1 : BOOL;
    Q2 : BOOL;
    Q3 : BOOL;
    CNT : INT;
    RUN : BOOL;
  END_VAR
  VAR
    r0 : DWORD;
    r1 : DWORD;
    r2 : DWORD;
    r3 : DWORD;
    rx : INT := 1;
  END_VAR

  (* check if number of runs is finished or rep = 0 which means continuous *)

  IF clk AND NOT rst THEN
  	run := (rep = 0) OR (rx <= rep);
  	IF run THEN
  		(* check for step counter reached and reset to 0 if cnt = steps *)
  		IF cnt = steps THEN
  			cnt := 0;
  		END_IF;

  		(* when cnt = 0 then reload the inputs into the registers *)
  		IF cnt = 0 THEN
  			r0 := in0;
  			r1 := in1;
  			r2 := in2;
  			r3 := in3;
  		END_IF;

  		(* when cnt < steps, shift the lowest bits to the outputs *)
  		IF (cnt < steps) THEN
              Q0 := BIT_OF_DWORD(r0,0); (* Q0 := r0.X0; *)
              Q1 := BIT_OF_DWORD(r1,0); (* Q1 := r1.X0; *)
              Q2 := BIT_OF_DWORD(r2,0); (* Q2 := r2.X0; *)
              Q3 := BIT_OF_DWORD(r3,0); (* Q3 := r3.X0; *)
  			r0 := SHR(r0,2); (* MUTATED: CONST_VALUE_REPLACE *)
  			r1 := SHR(r1,1);
  			r2 := SHR(r2,1);
  			r3 := SHR(r3,1);
  		END_IF;

  		(* increment the step counter *)
  		cnt := cnt +1;
  		IF (cnt = steps) AND (rep <> 0) THEN rx := rx +1; END_IF;
  		IF (rx > rep) AND (rep <> 0) THEN run := FALSE; END_IF;
  	END_IF;
  ELSE
  	IF rst THEN
  		run := FALSE;
  		Q0 := FALSE;
  		Q1 := FALSE;
  		Q2 := FALSE;
  		Q3 := FALSE;
  		r0 := DWORD#0;
  		r1 := DWORD#0;
  		r2 := DWORD#0;
  		r3 := DWORD#0;
  		cnt := 0;
  		rx := 1;
  	END_IF;
  END_IF;

  (*From OSCAT Library, www.oscat.de *)
END_FUNCTION_BLOCK

(* ---- M037.st ---- *)
FUNCTION_BLOCK GEN_BIT
  VAR_INPUT
    IN0 : DWORD;
    IN1 : DWORD;
    IN2 : DWORD;
    IN3 : DWORD;
    CLK : BOOL;
    STEPS : INT;
    REP : INT;
    RST : BOOL;
  END_VAR
  VAR_OUTPUT
    Q0 : BOOL;
    Q1 : BOOL;
    Q2 : BOOL;
    Q3 : BOOL;
    CNT : INT;
    RUN : BOOL;
  END_VAR
  VAR
    r0 : DWORD;
    r1 : DWORD;
    r2 : DWORD;
    r3 : DWORD;
    rx : INT := 1;
  END_VAR

  (* check if number of runs is finished or rep = 0 which means continuous *)

  IF clk AND NOT rst THEN
  	run := (rep = 0) OR (rx <= rep);
  	IF run THEN
  		(* check for step counter reached and reset to 0 if cnt = steps *)
  		IF cnt = steps THEN
  			cnt := 0;
  		END_IF;

  		(* when cnt = 0 then reload the inputs into the registers *)
  		IF cnt = 0 THEN
  			r0 := in0;
  			r1 := in1;
  			r2 := in2;
  			r3 := in3;
  		END_IF;

  		(* when cnt < steps, shift the lowest bits to the outputs *)
  		IF (cnt < steps) THEN
              Q0 := BIT_OF_DWORD(r0,0); (* Q0 := r0.X0; *)
              Q1 := BIT_OF_DWORD(r1,0); (* Q1 := r1.X0; *)
              Q2 := BIT_OF_DWORD(r2,0); (* Q2 := r2.X0; *)
              Q3 := BIT_OF_DWORD(r3,0); (* Q3 := r3.X0; *)
  			r0 := SHR(r0,1);
  			r1 := SHR(r1,2); (* MUTATED: CONST_VALUE_REPLACE *)
  			r2 := SHR(r2,1);
  			r3 := SHR(r3,1);
  		END_IF;

  		(* increment the step counter *)
  		cnt := cnt +1;
  		IF (cnt = steps) AND (rep <> 0) THEN rx := rx +1; END_IF;
  		IF (rx > rep) AND (rep <> 0) THEN run := FALSE; END_IF;
  	END_IF;
  ELSE
  	IF rst THEN
  		run := FALSE;
  		Q0 := FALSE;
  		Q1 := FALSE;
  		Q2 := FALSE;
  		Q3 := FALSE;
  		r0 := DWORD#0;
  		r1 := DWORD#0;
  		r2 := DWORD#0;
  		r3 := DWORD#0;
  		cnt := 0;
  		rx := 1;
  	END_IF;
  END_IF;

  (*From OSCAT Library, www.oscat.de *)
END_FUNCTION_BLOCK

(* ---- M038.st ---- *)
FUNCTION_BLOCK GEN_BIT
  VAR_INPUT
    IN0 : DWORD;
    IN1 : DWORD;
    IN2 : DWORD;
    IN3 : DWORD;
    CLK : BOOL;
    STEPS : INT;
    REP : INT;
    RST : BOOL;
  END_VAR
  VAR_OUTPUT
    Q0 : BOOL;
    Q1 : BOOL;
    Q2 : BOOL;
    Q3 : BOOL;
    CNT : INT;
    RUN : BOOL;
  END_VAR
  VAR
    r0 : DWORD;
    r1 : DWORD;
    r2 : DWORD;
    r3 : DWORD;
    rx : INT := 1;
  END_VAR

  (* check if number of runs is finished or rep = 0 which means continuous *)

  IF clk AND NOT rst THEN
  	run := (rep = 0) OR (rx <= rep);
  	IF run THEN
  		(* check for step counter reached and reset to 0 if cnt = steps *)
  		IF cnt = steps THEN
  			cnt := 0;
  		END_IF;

  		(* when cnt = 0 then reload the inputs into the registers *)
  		IF cnt = 0 THEN
  			r0 := in0;
  			r1 := in1;
  			r2 := in2;
  			r3 := in3;
  		END_IF;

  		(* when cnt < steps, shift the lowest bits to the outputs *)
  		IF (cnt < steps) THEN
              Q0 := BIT_OF_DWORD(r0,0); (* Q0 := r0.X0; *)
              Q1 := BIT_OF_DWORD(r1,0); (* Q1 := r1.X0; *)
              Q2 := BIT_OF_DWORD(r2,0); (* Q2 := r2.X0; *)
              Q3 := BIT_OF_DWORD(r3,0); (* Q3 := r3.X0; *)
  			r0 := SHR(r0,1);
  			r1 := SHR(r1,1);
  			r2 := SHR(r2,2); (* MUTATED: CONST_VALUE_REPLACE *)
  			r3 := SHR(r3,1);
  		END_IF;

  		(* increment the step counter *)
  		cnt := cnt +1;
  		IF (cnt = steps) AND (rep <> 0) THEN rx := rx +1; END_IF;
  		IF (rx > rep) AND (rep <> 0) THEN run := FALSE; END_IF;
  	END_IF;
  ELSE
  	IF rst THEN
  		run := FALSE;
  		Q0 := FALSE;
  		Q1 := FALSE;
  		Q2 := FALSE;
  		Q3 := FALSE;
  		r0 := DWORD#0;
  		r1 := DWORD#0;
  		r2 := DWORD#0;
  		r3 := DWORD#0;
  		cnt := 0;
  		rx := 1;
  	END_IF;
  END_IF;

  (*From OSCAT Library, www.oscat.de *)
END_FUNCTION_BLOCK

(* ---- M039.st ---- *)
FUNCTION_BLOCK GEN_BIT
  VAR_INPUT
    IN0 : DWORD;
    IN1 : DWORD;
    IN2 : DWORD;
    IN3 : DWORD;
    CLK : BOOL;
    STEPS : INT;
    REP : INT;
    RST : BOOL;
  END_VAR
  VAR_OUTPUT
    Q0 : BOOL;
    Q1 : BOOL;
    Q2 : BOOL;
    Q3 : BOOL;
    CNT : INT;
    RUN : BOOL;
  END_VAR
  VAR
    r0 : DWORD;
    r1 : DWORD;
    r2 : DWORD;
    r3 : DWORD;
    rx : INT := 1;
  END_VAR

  (* check if number of runs is finished or rep = 0 which means continuous *)

  IF clk AND NOT rst THEN
  	run := (rep = 0) OR (rx <= rep);
  	IF run THEN
  		(* check for step counter reached and reset to 0 if cnt = steps *)
  		IF cnt = steps THEN
  			cnt := 0;
  		END_IF;

  		(* when cnt = 0 then reload the inputs into the registers *)
  		IF cnt = 0 THEN
  			r0 := in0;
  			r1 := in1;
  			r2 := in2;
  			r3 := in3;
  		END_IF;

  		(* when cnt < steps, shift the lowest bits to the outputs *)
  		IF (cnt < steps) THEN
              Q0 := BIT_OF_DWORD(r0,0); (* Q0 := r0.X0; *)
              Q1 := BIT_OF_DWORD(r1,0); (* Q1 := r1.X0; *)
              Q2 := BIT_OF_DWORD(r2,0); (* Q2 := r2.X0; *)
              Q3 := BIT_OF_DWORD(r3,0); (* Q3 := r3.X0; *)
  			r0 := SHR(r0,1);
  			r1 := SHR(r1,1);
  			r2 := SHR(r2,1);
  			r3 := SHR(r3,2); (* MUTATED: CONST_VALUE_REPLACE *)
  		END_IF;

  		(* increment the step counter *)
  		cnt := cnt +1;
  		IF (cnt = steps) AND (rep <> 0) THEN rx := rx +1; END_IF;
  		IF (rx > rep) AND (rep <> 0) THEN run := FALSE; END_IF;
  	END_IF;
  ELSE
  	IF rst THEN
  		run := FALSE;
  		Q0 := FALSE;
  		Q1 := FALSE;
  		Q2 := FALSE;
  		Q3 := FALSE;
  		r0 := DWORD#0;
  		r1 := DWORD#0;
  		r2 := DWORD#0;
  		r3 := DWORD#0;
  		cnt := 0;
  		rx := 1;
  	END_IF;
  END_IF;

  (*From OSCAT Library, www.oscat.de *)
END_FUNCTION_BLOCK

(* ---- M040.st ---- *)
FUNCTION_BLOCK GEN_BIT
  VAR_INPUT
    IN0 : DWORD;
    IN1 : DWORD;
    IN2 : DWORD;
    IN3 : DWORD;
    CLK : BOOL;
    STEPS : INT;
    REP : INT;
    RST : BOOL;
  END_VAR
  VAR_OUTPUT
    Q0 : BOOL;
    Q1 : BOOL;
    Q2 : BOOL;
    Q3 : BOOL;
    CNT : INT;
    RUN : BOOL;
  END_VAR
  VAR
    r0 : DWORD;
    r1 : DWORD;
    r2 : DWORD;
    r3 : DWORD;
    rx : INT := 1;
  END_VAR

  (* check if number of runs is finished or rep = 0 which means continuous *)

  IF clk AND NOT rst THEN
  	run := (rep = 0) OR (rx <= rep);
  	IF run THEN
  		(* check for step counter reached and reset to 0 if cnt = steps *)
  		IF cnt = steps THEN
  			cnt := 0;
  		END_IF;

  		(* when cnt = 0 then reload the inputs into the registers *)
  		IF cnt = 0 THEN
  			r0 := in0;
  			r1 := in1;
  			r2 := in2;
  			r3 := in3;
  		END_IF;

  		(* when cnt < steps, shift the lowest bits to the outputs *)
  		IF (cnt < steps) THEN
              Q0 := BIT_OF_DWORD(r0,0); (* Q0 := r0.X0; *)
              Q1 := BIT_OF_DWORD(r1,0); (* Q1 := r1.X0; *)
              Q2 := BIT_OF_DWORD(r2,0); (* Q2 := r2.X0; *)
              Q3 := BIT_OF_DWORD(r3,0); (* Q3 := r3.X0; *)
  			r0 := SHR(r0,1);
  			r1 := SHR(r1,1);
  			r2 := SHR(r2,1);
  			r3 := SHR(r3,1);
  		END_IF;

  		(* increment the step counter *)
  		cnt := cnt +2; (* MUTATED: CONST_VALUE_REPLACE *)
  		IF (cnt = steps) AND (rep <> 0) THEN rx := rx +1; END_IF;
  		IF (rx > rep) AND (rep <> 0) THEN run := FALSE; END_IF;
  	END_IF;
  ELSE
  	IF rst THEN
  		run := FALSE;
  		Q0 := FALSE;
  		Q1 := FALSE;
  		Q2 := FALSE;
  		Q3 := FALSE;
  		r0 := DWORD#0;
  		r1 := DWORD#0;
  		r2 := DWORD#0;
  		r3 := DWORD#0;
  		cnt := 0;
  		rx := 1;
  	END_IF;
  END_IF;

  (*From OSCAT Library, www.oscat.de *)
END_FUNCTION_BLOCK

(* ---- M041.st ---- *)
FUNCTION_BLOCK GEN_BIT
  VAR_INPUT
    IN0 : DWORD;
    IN1 : DWORD;
    IN2 : DWORD;
    IN3 : DWORD;
    CLK : BOOL;
    STEPS : INT;
    REP : INT;
    RST : BOOL;
  END_VAR
  VAR_OUTPUT
    Q0 : BOOL;
    Q1 : BOOL;
    Q2 : BOOL;
    Q3 : BOOL;
    CNT : INT;
    RUN : BOOL;
  END_VAR
  VAR
    r0 : DWORD;
    r1 : DWORD;
    r2 : DWORD;
    r3 : DWORD;
    rx : INT := 1;
  END_VAR

  (* check if number of runs is finished or rep = 0 which means continuous *)

  IF clk AND NOT rst THEN
  	run := (rep = 0) OR (rx <= rep);
  	IF run THEN
  		(* check for step counter reached and reset to 0 if cnt = steps *)
  		IF cnt = steps THEN
  			cnt := 0;
  		END_IF;

  		(* when cnt = 0 then reload the inputs into the registers *)
  		IF cnt = 0 THEN
  			r0 := in0;
  			r1 := in1;
  			r2 := in2;
  			r3 := in3;
  		END_IF;

  		(* when cnt < steps, shift the lowest bits to the outputs *)
  		IF (cnt < steps) THEN
              Q0 := BIT_OF_DWORD(r0,0); (* Q0 := r0.X0; *)
              Q1 := BIT_OF_DWORD(r1,0); (* Q1 := r1.X0; *)
              Q2 := BIT_OF_DWORD(r2,0); (* Q2 := r2.X0; *)
              Q3 := BIT_OF_DWORD(r3,0); (* Q3 := r3.X0; *)
  			r0 := SHR(r0,1);
  			r1 := SHR(r1,1);
  			r2 := SHR(r2,1);
  			r3 := SHR(r3,1);
  		END_IF;

  		(* increment the step counter *)
  		cnt := cnt +1;
  		IF (cnt = steps) AND (rep <> 1) THEN rx := rx +1; END_IF; (* MUTATED: CONST_VALUE_REPLACE *)
  		IF (rx > rep) AND (rep <> 0) THEN run := FALSE; END_IF;
  	END_IF;
  ELSE
  	IF rst THEN
  		run := FALSE;
  		Q0 := FALSE;
  		Q1 := FALSE;
  		Q2 := FALSE;
  		Q3 := FALSE;
  		r0 := DWORD#0;
  		r1 := DWORD#0;
  		r2 := DWORD#0;
  		r3 := DWORD#0;
  		cnt := 0;
  		rx := 1;
  	END_IF;
  END_IF;

  (*From OSCAT Library, www.oscat.de *)
END_FUNCTION_BLOCK

(* ---- M042.st ---- *)
FUNCTION_BLOCK GEN_BIT
  VAR_INPUT
    IN0 : DWORD;
    IN1 : DWORD;
    IN2 : DWORD;
    IN3 : DWORD;
    CLK : BOOL;
    STEPS : INT;
    REP : INT;
    RST : BOOL;
  END_VAR
  VAR_OUTPUT
    Q0 : BOOL;
    Q1 : BOOL;
    Q2 : BOOL;
    Q3 : BOOL;
    CNT : INT;
    RUN : BOOL;
  END_VAR
  VAR
    r0 : DWORD;
    r1 : DWORD;
    r2 : DWORD;
    r3 : DWORD;
    rx : INT := 1;
  END_VAR

  (* check if number of runs is finished or rep = 0 which means continuous *)

  IF clk AND NOT rst THEN
  	run := (rep = 0) OR (rx <= rep);
  	IF run THEN
  		(* check for step counter reached and reset to 0 if cnt = steps *)
  		IF cnt = steps THEN
  			cnt := 0;
  		END_IF;

  		(* when cnt = 0 then reload the inputs into the registers *)
  		IF cnt = 0 THEN
  			r0 := in0;
  			r1 := in1;
  			r2 := in2;
  			r3 := in3;
  		END_IF;

  		(* when cnt < steps, shift the lowest bits to the outputs *)
  		IF (cnt < steps) THEN
              Q0 := BIT_OF_DWORD(r0,0); (* Q0 := r0.X0; *)
              Q1 := BIT_OF_DWORD(r1,0); (* Q1 := r1.X0; *)
              Q2 := BIT_OF_DWORD(r2,0); (* Q2 := r2.X0; *)
              Q3 := BIT_OF_DWORD(r3,0); (* Q3 := r3.X0; *)
  			r0 := SHR(r0,1);
  			r1 := SHR(r1,1);
  			r2 := SHR(r2,1);
  			r3 := SHR(r3,1);
  		END_IF;

  		(* increment the step counter *)
  		cnt := cnt +1;
  		IF (cnt = steps) AND (rep <> 0) THEN rx := rx +2; END_IF; (* MUTATED: CONST_VALUE_REPLACE *)
  		IF (rx > rep) AND (rep <> 0) THEN run := FALSE; END_IF;
  	END_IF;
  ELSE
  	IF rst THEN
  		run := FALSE;
  		Q0 := FALSE;
  		Q1 := FALSE;
  		Q2 := FALSE;
  		Q3 := FALSE;
  		r0 := DWORD#0;
  		r1 := DWORD#0;
  		r2 := DWORD#0;
  		r3 := DWORD#0;
  		cnt := 0;
  		rx := 1;
  	END_IF;
  END_IF;

  (*From OSCAT Library, www.oscat.de *)
END_FUNCTION_BLOCK

(* ---- M043.st ---- *)
FUNCTION_BLOCK GEN_BIT
  VAR_INPUT
    IN0 : DWORD;
    IN1 : DWORD;
    IN2 : DWORD;
    IN3 : DWORD;
    CLK : BOOL;
    STEPS : INT;
    REP : INT;
    RST : BOOL;
  END_VAR
  VAR_OUTPUT
    Q0 : BOOL;
    Q1 : BOOL;
    Q2 : BOOL;
    Q3 : BOOL;
    CNT : INT;
    RUN : BOOL;
  END_VAR
  VAR
    r0 : DWORD;
    r1 : DWORD;
    r2 : DWORD;
    r3 : DWORD;
    rx : INT := 1;
  END_VAR

  (* check if number of runs is finished or rep = 0 which means continuous *)

  IF clk AND NOT rst THEN
  	run := (rep = 0) OR (rx <= rep);
  	IF run THEN
  		(* check for step counter reached and reset to 0 if cnt = steps *)
  		IF cnt = steps THEN
  			cnt := 0;
  		END_IF;

  		(* when cnt = 0 then reload the inputs into the registers *)
  		IF cnt = 0 THEN
  			r0 := in0;
  			r1 := in1;
  			r2 := in2;
  			r3 := in3;
  		END_IF;

  		(* when cnt < steps, shift the lowest bits to the outputs *)
  		IF (cnt < steps) THEN
              Q0 := BIT_OF_DWORD(r0,0); (* Q0 := r0.X0; *)
              Q1 := BIT_OF_DWORD(r1,0); (* Q1 := r1.X0; *)
              Q2 := BIT_OF_DWORD(r2,0); (* Q2 := r2.X0; *)
              Q3 := BIT_OF_DWORD(r3,0); (* Q3 := r3.X0; *)
  			r0 := SHR(r0,1);
  			r1 := SHR(r1,1);
  			r2 := SHR(r2,1);
  			r3 := SHR(r3,1);
  		END_IF;

  		(* increment the step counter *)
  		cnt := cnt +1;
  		IF (cnt = steps) AND (rep <> 0) THEN rx := rx +1; END_IF;
  		IF (rx > rep) AND (rep <> 1) THEN run := FALSE; END_IF; (* MUTATED: CONST_VALUE_REPLACE *)
  	END_IF;
  ELSE
  	IF rst THEN
  		run := FALSE;
  		Q0 := FALSE;
  		Q1 := FALSE;
  		Q2 := FALSE;
  		Q3 := FALSE;
  		r0 := DWORD#0;
  		r1 := DWORD#0;
  		r2 := DWORD#0;
  		r3 := DWORD#0;
  		cnt := 0;
  		rx := 1;
  	END_IF;
  END_IF;

  (*From OSCAT Library, www.oscat.de *)
END_FUNCTION_BLOCK

(* ---- M044.st ---- *)
FUNCTION_BLOCK GEN_BIT
  VAR_INPUT
    IN0 : DWORD;
    IN1 : DWORD;
    IN2 : DWORD;
    IN3 : DWORD;
    CLK : BOOL;
    STEPS : INT;
    REP : INT;
    RST : BOOL;
  END_VAR
  VAR_OUTPUT
    Q0 : BOOL;
    Q1 : BOOL;
    Q2 : BOOL;
    Q3 : BOOL;
    CNT : INT;
    RUN : BOOL;
  END_VAR
  VAR
    r0 : DWORD;
    r1 : DWORD;
    r2 : DWORD;
    r3 : DWORD;
    rx : INT := 1;
  END_VAR

  (* check if number of runs is finished or rep = 0 which means continuous *)

  IF clk AND NOT rst THEN
  	run := (rep = 0) OR (rx <= rep);
  	IF run THEN
  		(* check for step counter reached and reset to 0 if cnt = steps *)
  		IF cnt = steps THEN
  			cnt := 0;
  		END_IF;

  		(* when cnt = 0 then reload the inputs into the registers *)
  		IF cnt = 0 THEN
  			r0 := in0;
  			r1 := in1;
  			r2 := in2;
  			r3 := in3;
  		END_IF;

  		(* when cnt < steps, shift the lowest bits to the outputs *)
  		IF (cnt < steps) THEN
              Q0 := BIT_OF_DWORD(r0,0); (* Q0 := r0.X0; *)
              Q1 := BIT_OF_DWORD(r1,0); (* Q1 := r1.X0; *)
              Q2 := BIT_OF_DWORD(r2,0); (* Q2 := r2.X0; *)
              Q3 := BIT_OF_DWORD(r3,0); (* Q3 := r3.X0; *)
  			r0 := SHR(r0,1);
  			r1 := SHR(r1,1);
  			r2 := SHR(r2,1);
  			r3 := SHR(r3,1);
  		END_IF;

  		(* increment the step counter *)
  		cnt := cnt +1;
  		IF (cnt = steps) AND (rep <> 0) THEN rx := rx +1; END_IF;
  		IF (rx > rep) AND (rep <> 0) THEN run := FALSE; END_IF;
  	END_IF;
  ELSE
  	IF rst THEN
  		run := FALSE;
  		Q0 := FALSE;
  		Q1 := FALSE;
  		Q2 := FALSE;
  		Q3 := FALSE;
  		r0 := DWORD#0;
  		r1 := DWORD#0;
  		r2 := DWORD#0;
  		r3 := DWORD#0;
  		cnt := 1; (* MUTATED: CONST_VALUE_REPLACE *)
  		rx := 1;
  	END_IF;
  END_IF;

  (*From OSCAT Library, www.oscat.de *)
END_FUNCTION_BLOCK

(* ---- M045.st ---- *)
FUNCTION_BLOCK GEN_BIT
  VAR_INPUT
    IN0 : DWORD;
    IN1 : DWORD;
    IN2 : DWORD;
    IN3 : DWORD;
    CLK : BOOL;
    STEPS : INT;
    REP : INT;
    RST : BOOL;
  END_VAR
  VAR_OUTPUT
    Q0 : BOOL;
    Q1 : BOOL;
    Q2 : BOOL;
    Q3 : BOOL;
    CNT : INT;
    RUN : BOOL;
  END_VAR
  VAR
    r0 : DWORD;
    r1 : DWORD;
    r2 : DWORD;
    r3 : DWORD;
    rx : INT := 1;
  END_VAR

  (* check if number of runs is finished or rep = 0 which means continuous *)

  IF clk AND NOT rst THEN
  	run := (rep = 0) OR (rx <= rep);
  	IF run THEN
  		(* check for step counter reached and reset to 0 if cnt = steps *)
  		IF cnt = steps THEN
  			cnt := 0;
  		END_IF;

  		(* when cnt = 0 then reload the inputs into the registers *)
  		IF cnt = 0 THEN
  			r0 := in0;
  			r1 := in1;
  			r2 := in2;
  			r3 := in3;
  		END_IF;

  		(* when cnt < steps, shift the lowest bits to the outputs *)
  		IF (cnt < steps) THEN
              Q0 := BIT_OF_DWORD(r0,0); (* Q0 := r0.X0; *)
              Q1 := BIT_OF_DWORD(r1,0); (* Q1 := r1.X0; *)
              Q2 := BIT_OF_DWORD(r2,0); (* Q2 := r2.X0; *)
              Q3 := BIT_OF_DWORD(r3,0); (* Q3 := r3.X0; *)
  			r0 := SHR(r0,1);
  			r1 := SHR(r1,1);
  			r2 := SHR(r2,1);
  			r3 := SHR(r3,1);
  		END_IF;

  		(* increment the step counter *)
  		cnt := cnt +1;
  		IF (cnt = steps) AND (rep <> 0) THEN rx := rx +1; END_IF;
  		IF (rx > rep) AND (rep <> 0) THEN run := FALSE; END_IF;
  	END_IF;
  ELSE
  	IF rst THEN
  		run := FALSE;
  		Q0 := FALSE;
  		Q1 := FALSE;
  		Q2 := FALSE;
  		Q3 := FALSE;
  		r0 := DWORD#0;
  		r1 := DWORD#0;
  		r2 := DWORD#0;
  		r3 := DWORD#0;
  		cnt := 0;
  		rx := 2; (* MUTATED: CONST_VALUE_REPLACE *)
  	END_IF;
  END_IF;

  (*From OSCAT Library, www.oscat.de *)
END_FUNCTION_BLOCK

(* ---- M046.st ---- *)
FUNCTION_BLOCK GEN_BIT
  VAR_INPUT
    IN0 : DWORD;
    IN1 : DWORD;
    IN2 : DWORD;
    IN3 : DWORD;
    CLK : BOOL;
    STEPS : INT;
    REP : INT;
    RST : BOOL;
  END_VAR
  VAR_OUTPUT
    Q0 : BOOL;
    Q1 : BOOL;
    Q2 : BOOL;
    Q3 : BOOL;
    CNT : INT;
    RUN : BOOL;
  END_VAR
  VAR
    r0 : DWORD;
    r1 : DWORD;
    r2 : DWORD;
    r3 : DWORD;
    rx : INT := 1;
  END_VAR

  (* check if number of runs is finished or rep = 0 which means continuous *)

  IF clk AND NOT rst THEN
  	run := (rep = 0) OR (rx <= rep);
  	IF run THEN
  		(* check for step counter reached and reset to 0 if cnt = steps *)
  		IF cnt = steps THEN
  			cnt := 0;
  		END_IF;

  		(* when cnt = 0 then reload the inputs into the registers *)
  		IF cnt = 0 THEN
  			r0 := in0;
  			r1 := in1;
  			r2 := in2;
  			r3 := in3;
  		END_IF;

  		(* when cnt < steps, shift the lowest bits to the outputs *)
  		IF (cnt < steps) THEN
              Q1 := BIT_OF_DWORD(r0,0); (* Q0 := r0.X0; *) (* MUTATED: VAR_REPLACE *)
              Q1 := BIT_OF_DWORD(r1,0); (* Q1 := r1.X0; *)
              Q2 := BIT_OF_DWORD(r2,0); (* Q2 := r2.X0; *)
              Q3 := BIT_OF_DWORD(r3,0); (* Q3 := r3.X0; *)
  			r0 := SHR(r0,1);
  			r1 := SHR(r1,1);
  			r2 := SHR(r2,1);
  			r3 := SHR(r3,1);
  		END_IF;

  		(* increment the step counter *)
  		cnt := cnt +1;
  		IF (cnt = steps) AND (rep <> 0) THEN rx := rx +1; END_IF;
  		IF (rx > rep) AND (rep <> 0) THEN run := FALSE; END_IF;
  	END_IF;
  ELSE
  	IF rst THEN
  		run := FALSE;
  		Q0 := FALSE;
  		Q1 := FALSE;
  		Q2 := FALSE;
  		Q3 := FALSE;
  		r0 := DWORD#0;
  		r1 := DWORD#0;
  		r2 := DWORD#0;
  		r3 := DWORD#0;
  		cnt := 0;
  		rx := 1;
  	END_IF;
  END_IF;

  (*From OSCAT Library, www.oscat.de *)
END_FUNCTION_BLOCK

(* ---- M047.st ---- *)
FUNCTION_BLOCK GEN_BIT
  VAR_INPUT
    IN0 : DWORD;
    IN1 : DWORD;
    IN2 : DWORD;
    IN3 : DWORD;
    CLK : BOOL;
    STEPS : INT;
    REP : INT;
    RST : BOOL;
  END_VAR
  VAR_OUTPUT
    Q0 : BOOL;
    Q1 : BOOL;
    Q2 : BOOL;
    Q3 : BOOL;
    CNT : INT;
    RUN : BOOL;
  END_VAR
  VAR
    r0 : DWORD;
    r1 : DWORD;
    r2 : DWORD;
    r3 : DWORD;
    rx : INT := 1;
  END_VAR

  (* check if number of runs is finished or rep = 0 which means continuous *)

  IF clk AND NOT rst THEN
  	run := (rep = 0) OR (rx <= rep);
  	IF run THEN
  		(* check for step counter reached and reset to 0 if cnt = steps *)
  		IF cnt = steps THEN
  			cnt := 0;
  		END_IF;

  		(* when cnt = 0 then reload the inputs into the registers *)
  		IF cnt = 0 THEN
  			r0 := in0;
  			r1 := in1;
  			r2 := in2;
  			r3 := in3;
  		END_IF;

  		(* when cnt < steps, shift the lowest bits to the outputs *)
  		IF (cnt < steps) THEN
              Q0 := BIT_OF_DWORD(r0,0); (* Q0 := r0.X0; *)
              Q2 := BIT_OF_DWORD(r1,0); (* Q1 := r1.X0; *) (* MUTATED: VAR_REPLACE *)
              Q2 := BIT_OF_DWORD(r2,0); (* Q2 := r2.X0; *)
              Q3 := BIT_OF_DWORD(r3,0); (* Q3 := r3.X0; *)
  			r0 := SHR(r0,1);
  			r1 := SHR(r1,1);
  			r2 := SHR(r2,1);
  			r3 := SHR(r3,1);
  		END_IF;

  		(* increment the step counter *)
  		cnt := cnt +1;
  		IF (cnt = steps) AND (rep <> 0) THEN rx := rx +1; END_IF;
  		IF (rx > rep) AND (rep <> 0) THEN run := FALSE; END_IF;
  	END_IF;
  ELSE
  	IF rst THEN
  		run := FALSE;
  		Q0 := FALSE;
  		Q1 := FALSE;
  		Q2 := FALSE;
  		Q3 := FALSE;
  		r0 := DWORD#0;
  		r1 := DWORD#0;
  		r2 := DWORD#0;
  		r3 := DWORD#0;
  		cnt := 0;
  		rx := 1;
  	END_IF;
  END_IF;

  (*From OSCAT Library, www.oscat.de *)
END_FUNCTION_BLOCK

(* ---- M048.st ---- *)
FUNCTION_BLOCK GEN_BIT
  VAR_INPUT
    IN0 : DWORD;
    IN1 : DWORD;
    IN2 : DWORD;
    IN3 : DWORD;
    CLK : BOOL;
    STEPS : INT;
    REP : INT;
    RST : BOOL;
  END_VAR
  VAR_OUTPUT
    Q0 : BOOL;
    Q1 : BOOL;
    Q2 : BOOL;
    Q3 : BOOL;
    CNT : INT;
    RUN : BOOL;
  END_VAR
  VAR
    r0 : DWORD;
    r1 : DWORD;
    r2 : DWORD;
    r3 : DWORD;
    rx : INT := 1;
  END_VAR

  (* check if number of runs is finished or rep = 0 which means continuous *)

  IF clk AND NOT rst THEN
  	run := (rep = 0) OR (rx <= rep);
  	IF run THEN
  		(* check for step counter reached and reset to 0 if cnt = steps *)
  		IF cnt = steps THEN
  			cnt := 0;
  		END_IF;

  		(* when cnt = 0 then reload the inputs into the registers *)
  		IF cnt = 0 THEN
  			r0 := in0;
  			r1 := in1;
  			r2 := in2;
  			r3 := in3;
  		END_IF;

  		(* when cnt < steps, shift the lowest bits to the outputs *)
  		IF (cnt < steps) THEN
              Q0 := BIT_OF_DWORD(r0,0); (* Q0 := r0.X0; *)
              Q1 := BIT_OF_DWORD(r1,0); (* Q1 := r1.X0; *)
              Q3 := BIT_OF_DWORD(r2,0); (* Q2 := r2.X0; *) (* MUTATED: VAR_REPLACE *)
              Q3 := BIT_OF_DWORD(r3,0); (* Q3 := r3.X0; *)
  			r0 := SHR(r0,1);
  			r1 := SHR(r1,1);
  			r2 := SHR(r2,1);
  			r3 := SHR(r3,1);
  		END_IF;

  		(* increment the step counter *)
  		cnt := cnt +1;
  		IF (cnt = steps) AND (rep <> 0) THEN rx := rx +1; END_IF;
  		IF (rx > rep) AND (rep <> 0) THEN run := FALSE; END_IF;
  	END_IF;
  ELSE
  	IF rst THEN
  		run := FALSE;
  		Q0 := FALSE;
  		Q1 := FALSE;
  		Q2 := FALSE;
  		Q3 := FALSE;
  		r0 := DWORD#0;
  		r1 := DWORD#0;
  		r2 := DWORD#0;
  		r3 := DWORD#0;
  		cnt := 0;
  		rx := 1;
  	END_IF;
  END_IF;

  (*From OSCAT Library, www.oscat.de *)
END_FUNCTION_BLOCK

(* ---- M049.st ---- *)
FUNCTION_BLOCK GEN_BIT
  VAR_INPUT
    IN0 : DWORD;
    IN1 : DWORD;
    IN2 : DWORD;
    IN3 : DWORD;
    CLK : BOOL;
    STEPS : INT;
    REP : INT;
    RST : BOOL;
  END_VAR
  VAR_OUTPUT
    Q0 : BOOL;
    Q1 : BOOL;
    Q2 : BOOL;
    Q3 : BOOL;
    CNT : INT;
    RUN : BOOL;
  END_VAR
  VAR
    r0 : DWORD;
    r1 : DWORD;
    r2 : DWORD;
    r3 : DWORD;
    rx : INT := 1;
  END_VAR

  (* check if number of runs is finished or rep = 0 which means continuous *)

  IF clk AND NOT rst THEN
  	run := (rep = 0) OR (rx <= rep);
  	IF run THEN
  		(* check for step counter reached and reset to 0 if cnt = steps *)
  		IF cnt = steps THEN
  			cnt := 0;
  		END_IF;

  		(* when cnt = 0 then reload the inputs into the registers *)
  		IF cnt = 0 THEN
  			r0 := in0;
  			r1 := in1;
  			r2 := in2;
  			r3 := in3;
  		END_IF;

  		(* when cnt < steps, shift the lowest bits to the outputs *)
  		IF (cnt < steps) THEN
              Q0 := BIT_OF_DWORD(r0,0); (* Q0 := r0.X0; *)
              Q1 := BIT_OF_DWORD(r1,0); (* Q1 := r1.X0; *)
              Q2 := BIT_OF_DWORD(r2,0); (* Q2 := r2.X0; *)
              RUN := BIT_OF_DWORD(r3,0); (* Q3 := r3.X0; *) (* MUTATED: VAR_REPLACE *)
  			r0 := SHR(r0,1);
  			r1 := SHR(r1,1);
  			r2 := SHR(r2,1);
  			r3 := SHR(r3,1);
  		END_IF;

  		(* increment the step counter *)
  		cnt := cnt +1;
  		IF (cnt = steps) AND (rep <> 0) THEN rx := rx +1; END_IF;
  		IF (rx > rep) AND (rep <> 0) THEN run := FALSE; END_IF;
  	END_IF;
  ELSE
  	IF rst THEN
  		run := FALSE;
  		Q0 := FALSE;
  		Q1 := FALSE;
  		Q2 := FALSE;
  		Q3 := FALSE;
  		r0 := DWORD#0;
  		r1 := DWORD#0;
  		r2 := DWORD#0;
  		r3 := DWORD#0;
  		cnt := 0;
  		rx := 1;
  	END_IF;
  END_IF;

  (*From OSCAT Library, www.oscat.de *)
END_FUNCTION_BLOCK

(* ---- M050.st ---- *)
FUNCTION_BLOCK GEN_BIT
  VAR_INPUT
    IN0 : DWORD;
    IN1 : DWORD;
    IN2 : DWORD;
    IN3 : DWORD;
    CLK : BOOL;
    STEPS : INT;
    REP : INT;
    RST : BOOL;
  END_VAR
  VAR_OUTPUT
    Q0 : BOOL;
    Q1 : BOOL;
    Q2 : BOOL;
    Q3 : BOOL;
    CNT : INT;
    RUN : BOOL;
  END_VAR
  VAR
    r0 : DWORD;
    r1 : DWORD;
    r2 : DWORD;
    r3 : DWORD;
    rx : INT := 1;
  END_VAR

  (* check if number of runs is finished or rep = 0 which means continuous *)

  IF clk AND NOT rst THEN
  	run := (rep = 0) OR (rx <= rep);
  	IF run THEN
  		(* check for step counter reached and reset to 0 if cnt = steps *)
  		IF cnt = steps THEN
  			cnt := 0;
  		END_IF;

  		(* when cnt = 0 then reload the inputs into the registers *)
  		IF cnt = 0 THEN
  			r0 := in0;
  			r1 := in1;
  			r2 := in2;
  			r3 := in3;
  		END_IF;

  		(* when cnt < steps, shift the lowest bits to the outputs *)
  		IF (cnt < steps) THEN
              Q0 := NOT (BIT_OF_DWORD(r0,0)); (* Q0 := r0.X0; *) (* MUTATED: ASSIGN_NEGATE *)
              Q1 := BIT_OF_DWORD(r1,0); (* Q1 := r1.X0; *)
              Q2 := BIT_OF_DWORD(r2,0); (* Q2 := r2.X0; *)
              Q3 := BIT_OF_DWORD(r3,0); (* Q3 := r3.X0; *)
  			r0 := SHR(r0,1);
  			r1 := SHR(r1,1);
  			r2 := SHR(r2,1);
  			r3 := SHR(r3,1);
  		END_IF;

  		(* increment the step counter *)
  		cnt := cnt +1;
  		IF (cnt = steps) AND (rep <> 0) THEN rx := rx +1; END_IF;
  		IF (rx > rep) AND (rep <> 0) THEN run := FALSE; END_IF;
  	END_IF;
  ELSE
  	IF rst THEN
  		run := FALSE;
  		Q0 := FALSE;
  		Q1 := FALSE;
  		Q2 := FALSE;
  		Q3 := FALSE;
  		r0 := DWORD#0;
  		r1 := DWORD#0;
  		r2 := DWORD#0;
  		r3 := DWORD#0;
  		cnt := 0;
  		rx := 1;
  	END_IF;
  END_IF;

  (*From OSCAT Library, www.oscat.de *)
END_FUNCTION_BLOCK

(* ---- M051.st ---- *)
FUNCTION_BLOCK GEN_BIT
  VAR_INPUT
    IN0 : DWORD;
    IN1 : DWORD;
    IN2 : DWORD;
    IN3 : DWORD;
    CLK : BOOL;
    STEPS : INT;
    REP : INT;
    RST : BOOL;
  END_VAR
  VAR_OUTPUT
    Q0 : BOOL;
    Q1 : BOOL;
    Q2 : BOOL;
    Q3 : BOOL;
    CNT : INT;
    RUN : BOOL;
  END_VAR
  VAR
    r0 : DWORD;
    r1 : DWORD;
    r2 : DWORD;
    r3 : DWORD;
    rx : INT := 1;
  END_VAR

  (* check if number of runs is finished or rep = 0 which means continuous *)

  IF clk AND NOT rst THEN
  	run := (rep = 0) OR (rx <= rep);
  	IF run THEN
  		(* check for step counter reached and reset to 0 if cnt = steps *)
  		IF cnt = steps THEN
  			cnt := 0;
  		END_IF;

  		(* when cnt = 0 then reload the inputs into the registers *)
  		IF cnt = 0 THEN
  			r0 := in0;
  			r1 := in1;
  			r2 := in2;
  			r3 := in3;
  		END_IF;

  		(* when cnt < steps, shift the lowest bits to the outputs *)
  		IF (cnt < steps) THEN
              Q0 := BIT_OF_DWORD(r0,0); (* Q0 := NOT (r0.X0); *) (* MUTATED: ASSIGN_NEGATE *)
              Q1 := BIT_OF_DWORD(r1,0); (* Q1 := r1.X0; *)
              Q2 := BIT_OF_DWORD(r2,0); (* Q2 := r2.X0; *)
              Q3 := BIT_OF_DWORD(r3,0); (* Q3 := r3.X0; *)
  			r0 := SHR(r0,1);
  			r1 := SHR(r1,1);
  			r2 := SHR(r2,1);
  			r3 := SHR(r3,1);
  		END_IF;

  		(* increment the step counter *)
  		cnt := cnt +1;
  		IF (cnt = steps) AND (rep <> 0) THEN rx := rx +1; END_IF;
  		IF (rx > rep) AND (rep <> 0) THEN run := FALSE; END_IF;
  	END_IF;
  ELSE
  	IF rst THEN
  		run := FALSE;
  		Q0 := FALSE;
  		Q1 := FALSE;
  		Q2 := FALSE;
  		Q3 := FALSE;
  		r0 := DWORD#0;
  		r1 := DWORD#0;
  		r2 := DWORD#0;
  		r3 := DWORD#0;
  		cnt := 0;
  		rx := 1;
  	END_IF;
  END_IF;

  (*From OSCAT Library, www.oscat.de *)
END_FUNCTION_BLOCK

(* ---- M052.st ---- *)
FUNCTION_BLOCK GEN_BIT
  VAR_INPUT
    IN0 : DWORD;
    IN1 : DWORD;
    IN2 : DWORD;
    IN3 : DWORD;
    CLK : BOOL;
    STEPS : INT;
    REP : INT;
    RST : BOOL;
  END_VAR
  VAR_OUTPUT
    Q0 : BOOL;
    Q1 : BOOL;
    Q2 : BOOL;
    Q3 : BOOL;
    CNT : INT;
    RUN : BOOL;
  END_VAR
  VAR
    r0 : DWORD;
    r1 : DWORD;
    r2 : DWORD;
    r3 : DWORD;
    rx : INT := 1;
  END_VAR

  (* check if number of runs is finished or rep = 0 which means continuous *)

  IF clk AND NOT rst THEN
  	run := (rep = 0) OR (rx <= rep);
  	IF run THEN
  		(* check for step counter reached and reset to 0 if cnt = steps *)
  		IF cnt = steps THEN
  			cnt := 0;
  		END_IF;

  		(* when cnt = 0 then reload the inputs into the registers *)
  		IF cnt = 0 THEN
  			r0 := in0;
  			r1 := in1;
  			r2 := in2;
  			r3 := in3;
  		END_IF;

  		(* when cnt < steps, shift the lowest bits to the outputs *)
  		IF (cnt < steps) THEN
              Q0 := BIT_OF_DWORD(r0,0); (* Q0 := r0.X0; *)
              Q1 := NOT (BIT_OF_DWORD(r1,0)); (* Q1 := r1.X0; *) (* MUTATED: ASSIGN_NEGATE *)
              Q2 := BIT_OF_DWORD(r2,0); (* Q2 := r2.X0; *)
              Q3 := BIT_OF_DWORD(r3,0); (* Q3 := r3.X0; *)
  			r0 := SHR(r0,1);
  			r1 := SHR(r1,1);
  			r2 := SHR(r2,1);
  			r3 := SHR(r3,1);
  		END_IF;

  		(* increment the step counter *)
  		cnt := cnt +1;
  		IF (cnt = steps) AND (rep <> 0) THEN rx := rx +1; END_IF;
  		IF (rx > rep) AND (rep <> 0) THEN run := FALSE; END_IF;
  	END_IF;
  ELSE
  	IF rst THEN
  		run := FALSE;
  		Q0 := FALSE;
  		Q1 := FALSE;
  		Q2 := FALSE;
  		Q3 := FALSE;
  		r0 := DWORD#0;
  		r1 := DWORD#0;
  		r2 := DWORD#0;
  		r3 := DWORD#0;
  		cnt := 0;
  		rx := 1;
  	END_IF;
  END_IF;

  (*From OSCAT Library, www.oscat.de *)
END_FUNCTION_BLOCK
